(* IEC 61131-3 sources: plc-st-coding-agent/progress/evidence/f14_v6_public_pilot_20261112/jobs/codex_minimax-m27, 42 files *)

(* ---- public-easy-01.candidate_01.st ---- *)
(*
ENGINEERING_CONTRACT
================================================================================
State Machine: Automated Filling Line (5-stage sequential + reset)
Clause ID | Output/State    | Activation          | Retention       | Reset
----------|-----------------|---------------------|-----------------|------------------
PUB003    | Pump_Motor      | bottleSensor=1      | Hold in CLEANING| cleaningConfirmButton (→FILLING)
PUB004    | Filling_Valve   | cleaningConfirmBtn  | Hold in FILLING | fillingConfirmButton (→CAPPING)
PUB005    | Capping_Machine | fillingConfirmBtn   | Hold in CAPPING | cappingConfirmButton (→PACKING)
PUB006    | Packing_Machine | cappingConfirmBtn   | Hold in PACKING | packingConfirmButton (→COMPLETE)
PUB007    | Completion_Light| packingConfirmBtn   | Hold until RESET| finishedButton (→IDLE)
PUB008    | (finishedButton)| Reset all, cycle end| N/A             | Automatic →IDLE
--------------------------------------------------------------------------------
Priority: Same-scan sequential (IDLE→CLEANING→FILLING→CAPPING→PACKING→COMPLETE→IDLE)
Units: None (binary signals, no timeouts specified)
Boundary: bottleSensor rising edge starts CLEANING; finishedButton resets COMPLETE→IDLE
--------------------------------------------------------------------------------
CONTRACT_RULES []
================================================================================
*)

FUNCTION_BLOCK FillingLineControl
VAR_INPUT
    bottleSensor          : BOOL;
    cleaningConfirmButton : BOOL;
    fillingConfirmButton  : BOOL;
    cappingConfirmButton  : BOOL;
    packingConfirmButton  : BOOL;
    finishedButton        : BOOL;
END_VAR
VAR_OUTPUT
    Pump_Motor      : BOOL;
    Filling_Valve   : BOOL;
    Capping_Machine : BOOL;
    Packing_Machine : BOOL;
    Completion_Light: BOOL;
END_VAR
VAR
    eState : INT;
END_VAR

// State enumeration: 0=IDLE, 1=CLEANING, 2=FILLING, 3=CAPPING, 4=PACKING, 5=COMPLETE
CASE eState OF
    0: // IDLE
        Pump_Motor       := FALSE;
        Filling_Valve    := FALSE;
        Capping_Machine  := FALSE;
        Packing_Machine  := FALSE;
        Completion_Light := FALSE;
        IF bottleSensor THEN
            eState := 1; // → CLEANING
        END_IF;

    1: // CLEANING
        Pump_Motor       := TRUE;
        Filling_Valve    := FALSE;
        Capping_Machine  := FALSE;
        Packing_Machine  := FALSE;
        Completion_Light := FALSE;
        IF cleaningConfirmButton THEN
            eState := 2; // → FILLING
        END_IF;

    2: // FILLING
        Pump_Motor       := FALSE;
        Filling_Valve    := TRUE;
        Capping_Machine  := FALSE;
        Packing_Machine  := FALSE;
        Completion_Light := FALSE;
        IF fillingConfirmButton THEN
            eState := 3; // → CAPPING
        END_IF;

    3: // CAPPING
        Pump_Motor       := FALSE;
        Filling_Valve    := FALSE;
        Capping_Machine  := TRUE;
        Packing_Machine  := FALSE;
        Completion_Light := FALSE;
        IF cappingConfirmButton THEN
            eState := 4; // → PACKING
        END_IF;

    4: // PACKING
        Pump_Motor       := FALSE;
        Filling_Valve    := FALSE;
        Capping_Machine  := FALSE;
        Packing_Machine  := TRUE;
        Completion_Light := FALSE;
        IF packingConfirmButton THEN
            eState := 5; // → COMPLETE
        END_IF;

    5: // COMPLETE
        Pump_Motor       := FALSE;
        Filling_Valve    := FALSE;
        Capping_Machine  := FALSE;
        Packing_Machine  := FALSE;
        Completion_Light := TRUE;
        IF finishedButton THEN
            eState := 0; // → IDLE (cycle reset)
        END_IF;

END_CASE;

END_FUNCTION_BLOCK

(* ---- public-easy-01.candidate_02.st ---- *)
(*
ENGINEERING_CONTRACT
================================================================================
State Machine: Automated Filling Line (5-stage sequential + reset)
Clause ID | Output/State    | Activation          | Retention       | Reset
----------|-----------------|---------------------|-----------------|------------------
PUB003    | Pump_Motor      | bottleSensor=1      | Hold in CLEANING| cleaningConfirmButton (→FILLING)
PUB004    | Filling_Valve   | cleaningConfirmBtn  | Hold in FILLING | fillingConfirmButton (→CAPPING)
PUB005    | Capping_Machine | fillingConfirmBtn   | Hold in CAPPING | cappingConfirmButton (→PACKING)
PUB006    | Packing_Machine | cappingConfirmBtn   | Hold in PACKING | packingConfirmButton (→COMPLETE)
PUB007    | Completion_Light| packingConfirmBtn   | Hold until RESET| finishedButton (→IDLE)
PUB008    | (finishedButton)| Reset all, cycle end| N/A             | Automatic →IDLE
--------------------------------------------------------------------------------
Priority: Same-scan sequential (IDLE→CLEANING→FILLING→CAPPING→PACKING→COMPLETE→IDLE)
Units: None (binary signals, no timeouts specified)
Boundary: bottleSensor rising edge starts CLEANING; finishedButton resets COMPLETE→IDLE
--------------------------------------------------------------------------------
CONTRACT_RULES []
================================================================================
*)

FUNCTION_BLOCK FillingLineControl
VAR_INPUT
    bottleSensor          : BOOL;
    cleaningConfirmButton : BOOL;
    fillingConfirmButton  : BOOL;
    cappingConfirmButton  : BOOL;
    packingConfirmButton  : BOOL;
    finishedButton        : BOOL;
END_VAR
VAR_OUTPUT
    Pump_Motor      : BOOL;
    Filling_Valve   : BOOL;
    Capping_Machine : BOOL;
    Packing_Machine : BOOL;
    Completion_Light: BOOL;
END_VAR
VAR
    eState : INT;
END_VAR

// State: 0=IDLE, 1=CLEANING, 2=FILLING, 3=CAPPING, 4=PACKING, 5=COMPLETE
// Multiple transitions within same scan when conditions allow
IF eState = 0 AND bottleSensor THEN
    eState := 1;
END_IF;

IF eState = 1 AND cleaningConfirmButton THEN
    eState := 2;
END_IF;

IF eState = 2 AND fillingConfirmButton THEN
    eState := 3;
END_IF;

IF eState = 3 AND cappingConfirmButton THEN
    eState := 4;
END_IF;

IF eState = 4 AND packingConfirmButton THEN
    eState := 5;
END_IF;

IF eState = 5 AND finishedButton THEN
    eState := 0;
END_IF;

// Output assignment based on current state
IF eState = 1 THEN
    Pump_Motor := TRUE;
END_IF;

IF eState = 2 THEN
    Filling_Valve := TRUE;
END_IF;

IF eState = 3 THEN
    Capping_Machine := TRUE;
END_IF;

IF eState = 4 THEN
    Packing_Machine := TRUE;
END_IF;

IF eState = 5 THEN
    Completion_Light := TRUE;
END_IF;

END_FUNCTION_BLOCK

(* ---- public-easy-01.candidate_03.st ---- *)
(*
ENGINEERING_CONTRACT
================================================================================
State Machine: Automated Filling Line (5-stage sequential + reset)
Clause ID | Output/State    | Activation          | Retention       | Reset
----------|-----------------|---------------------|-----------------|------------------
PUB003    | Pump_Motor      | bottleSensor=1      | Hold in CLEANING| cleaningConfirmButton (→FILLING)
PUB004    | Filling_Valve   | cleaningConfirmBtn  | Hold in FILLING | fillingConfirmButton (→CAPPING)
PUB005    | Capping_Machine | fillingConfirmBtn   | Hold in CAPPING | cappingConfirmButton (→PACKING)
PUB006    | Packing_Machine | cappingConfirmBtn   | Hold in PACKING | packingConfirmButton (→COMPLETE)
PUB007    | Completion_Light| packingConfirmBtn   | Hold until RESET| finishedButton (→IDLE)
PUB008    | (finishedButton)| Reset all, cycle end| N/A             | Automatic →IDLE
--------------------------------------------------------------------------------
Priority: Same-scan sequential (IDLE→CLEANING→FILLING→CAPPING→PACKING→COMPLETE→IDLE)
Units: None (binary signals, no timeouts specified)
Boundary: bottleSensor rising edge starts CLEANING; finishedButton resets COMPLETE→IDLE
--------------------------------------------------------------------------------
CONTRACT_RULES []
================================================================================
*)

FUNCTION_BLOCK FillingLineControl
VAR_INPUT
    bottleSensor          : BOOL;
    cleaningConfirmButton : BOOL;
    fillingConfirmButton  : BOOL;
    cappingConfirmButton  : BOOL;
    packingConfirmButton  : BOOL;
    finishedButton        : BOOL;
END_VAR
VAR_OUTPUT
    Pump_Motor      : BOOL;
    Filling_Valve   : BOOL;
    Capping_Machine : BOOL;
    Packing_Machine : BOOL;
    Completion_Light: BOOL;
END_VAR
VAR
    eState : INT;
END_VAR

// State: 0=IDLE, 1=CLEANING, 2=FILLING, 3=CAPPING, 4=PACKING, 5=COMPLETE
// Reset all outputs each scan to ensure clean state transitions
Pump_Motor      := FALSE;
Filling_Valve   := FALSE;
Capping_Machine := FALSE;
Packing_Machine := FALSE;
Completion_Light:= FALSE;

// State transitions - sequential same-scan processing
IF eState = 0 AND bottleSensor THEN
    eState := 1;
END_IF;

IF eState = 1 AND cleaningConfirmButton THEN
    eState := 2;
END_IF;

IF eState = 2 AND fillingConfirmButton THEN
    eState := 3;
END_IF;

IF eState = 3 AND cappingConfirmButton THEN
    eState := 4;
END_IF;

IF eState = 4 AND packingConfirmButton THEN
    eState := 5;
END_IF;

IF eState = 5 AND finishedButton THEN
    eState := 0;
END_IF;

// Output activation based on current state
IF eState = 1 THEN
    Pump_Motor := TRUE;
END_IF;

IF eState = 2 THEN
    Filling_Valve := TRUE;
END_IF;

IF eState = 3 THEN
    Capping_Machine := TRUE;
END_IF;

IF eState = 4 THEN
    Packing_Machine := TRUE;
END_IF;

IF eState = 5 THEN
    Completion_Light := TRUE;
END_IF;

END_FUNCTION_BLOCK

(* ---- public-easy-01.candidate_04.st ---- *)
Looking at the checkpoint, tc-08 shows ALL outputs TRUE when `finishedButton=true` from a prior state. The issue is that outputs never get reset when transitioning between states—they only get set TRUE but never set FALSE.

(*
ENGINEERING_CONTRACT
================================================================================
State Machine: Automated Filling Line (5-stage sequential + reset)
Clause ID | Output/State    | Activation          | Retention       | Reset
----------|-----------------|---------------------|-----------------|------------------
PUB003    | Pump_Motor      | bottleSensor=1      | Hold in CLEANING| Implicit (output cleared on state exit)
PUB004    | Filling_Valve   | cleaningConfirmBtn  | Hold in FILLING | Implicit (output cleared on state exit)
PUB005    | Capping_Machine | fillingConfirmBtn   | Hold in CAPPING | Implicit (output cleared on state exit)
PUB006    | Packing_Machine | cappingConfirmBtn   | Hold in PACKING | Implicit (output cleared on state exit)
PUB007    | Completion_Light| packingConfirmBtn   | Hold in COMPLETE| Implicit (output cleared on finishedButton reset)
PUB008    | (finishedButton)| Reset all outputs   | N/A             | Automatic →IDLE
--------------------------------------------------------------------------------
Priority: Same-scan sequential (IDLE→CLEANING→FILLING→CAPPING→PACKING→COMPLETE→IDLE)
Units: None (binary signals, no timeouts specified)
Boundary: Outputs are level-based; cleared when state exits, no edge-only behavior
--------------------------------------------------------------------------------
CONTRACT_RULES []
================================================================================
*)

FUNCTION_BLOCK FillingLineControl
VAR_INPUT
    bottleSensor          : BOOL;
    cleaningConfirmButton : BOOL;
    fillingConfirmButton  : BOOL;
    cappingConfirmButton  : BOOL;
    packingConfirmButton  : BOOL;
    finishedButton        : BOOL;
END_VAR
VAR_OUTPUT
    Pump_Motor      : BOOL;
    Filling_Valve   : BOOL;
    Capping_Machine : BOOL;
    Packing_Machine : BOOL;
    Completion_Light: BOOL;
END_VAR
VAR
    eState : INT;
END_VAR

// State: 0=IDLE, 1=CLEANING, 2=FILLING, 3=CAPPING, 4=PACKING, 5=COMPLETE
// Clear all outputs first (no latching across state transitions)
Pump_Motor      := FALSE;
Filling_Valve   := FALSE;
Capping_Machine := FALSE;
Packing_Machine := FALSE;
Completion_Light:= FALSE;

// State transitions (same-scan sequential)
IF eState = 0 AND bottleSensor THEN
    eState := 1;
END_IF;

IF eState = 1 AND cleaningConfirmButton THEN
    eState := 2;
END_IF;

IF eState = 2 AND fillingConfirmButton THEN
    eState := 3;
END_IF;

IF eState = 3 AND cappingConfirmButton THEN
    eState := 4;
END_IF;

IF eState = 4 AND packingConfirmButton THEN
    eState := 5;
END_IF;

IF eState = 5 AND finishedButton THEN
    eState := 0;
END_IF;

// Output assignment based on current state (level-based, cleared on exit)
IF eState = 1 THEN
    Pump_Motor := TRUE;
END_IF;

IF eState = 2 THEN
    Filling_Valve := TRUE;
END_IF;

IF eState = 3 THEN
    Capping_Machine := TRUE;
END_IF;

IF eState = 4 THEN
    Packing_Machine := TRUE;
END_IF;

IF eState = 5 THEN
    Completion_Light := TRUE;
END_IF;

END_FUNCTION_BLOCK

(* ---- public-easy-01.raw_candidate_01.st ---- *)
(*
ENGINEERING_CONTRACT
================================================================================
State Machine: Automated Filling Line (5-stage sequential + reset)
Clause ID | Output/State    | Activation          | Retention       | Reset
----------|-----------------|---------------------|-----------------|------------------
PUB003    | Pump_Motor      | bottleSensor=1      | Hold in CLEANING| cleaningConfirmButton (→FILLING)
PUB004    | Filling_Valve   | cleaningConfirmBtn  | Hold in FILLING | fillingConfirmButton (→CAPPING)
PUB005    | Capping_Machine | fillingConfirmBtn   | Hold in CAPPING | cappingConfirmButton (→PACKING)
PUB006    | Packing_Machine | cappingConfirmBtn   | Hold in PACKING | packingConfirmButton (→COMPLETE)
PUB007    | Completion_Light| packingConfirmBtn   | Hold until RESET| finishedButton (→IDLE)
PUB008    | (finishedButton)| Reset all, cycle end| N/A             | Automatic →IDLE
--------------------------------------------------------------------------------
Priority: Same-scan sequential (IDLE→CLEANING→FILLING→CAPPING→PACKING→COMPLETE→IDLE)
Units: None (binary signals, no timeouts specified)
Boundary: bottleSensor rising edge starts CLEANING; finishedButton resets COMPLETE→IDLE
--------------------------------------------------------------------------------
CONTRACT_RULES []
================================================================================
*)

FUNCTION_BLOCK FillingLineControl
VAR_INPUT
    bottleSensor          : BOOL;
    cleaningConfirmButton : BOOL;
    fillingConfirmButton  : BOOL;
    cappingConfirmButton  : BOOL;
    packingConfirmButton  : BOOL;
    finishedButton        : BOOL;
END_VAR
VAR_OUTPUT
    Pump_Motor      : BOOL;
    Filling_Valve   : BOOL;
    Capping_Machine : BOOL;
    Packing_Machine : BOOL;
    Completion_Light: BOOL;
END_VAR
VAR
    eState : INT;
END_VAR

// State enumeration: 0=IDLE, 1=CLEANING, 2=FILLING, 3=CAPPING, 4=PACKING, 5=COMPLETE
CASE eState OF
    0: // IDLE
        Pump_Motor       := FALSE;
        Filling_Valve    := FALSE;
        Capping_Machine  := FALSE;
        Packing_Machine  := FALSE;
        Completion_Light := FALSE;
        IF bottleSensor THEN
            eState := 1; // → CLEANING
        END_IF;

    1: // CLEANING
        Pump_Motor       := TRUE;
        Filling_Valve    := FALSE;
        Capping_Machine  := FALSE;
        Packing_Machine  := FALSE;
        Completion_Light := FALSE;
        IF cleaningConfirmButton THEN
            eState := 2; // → FILLING
        END_IF;

    2: // FILLING
        Pump_Motor       := FALSE;
        Filling_Valve    := TRUE;
        Capping_Machine  := FALSE;
        Packing_Machine  := FALSE;
        Completion_Light := FALSE;
        IF fillingConfirmButton THEN
            eState := 3; // → CAPPING
        END_IF;

    3: // CAPPING
        Pump_Motor       := FALSE;
        Filling_Valve    := FALSE;
        Capping_Machine  := TRUE;
        Packing_Machine  := FALSE;
        Completion_Light := FALSE;
        IF cappingConfirmButton THEN
            eState := 4; // → PACKING
        END_IF;

    4: // PACKING
        Pump_Motor       := FALSE;
        Filling_Valve    := FALSE;
        Capping_Machine  := FALSE;
        Packing_Machine  := TRUE;
        Completion_Light := FALSE;
        IF packingConfirmButton THEN
            eState := 5; // → COMPLETE
        END_IF;

    5: // COMPLETE
        Pump_Motor       := FALSE;
        Filling_Valve    := FALSE;
        Capping_Machine  := FALSE;
        Packing_Machine  := FALSE;
        Completion_Light := TRUE;
        IF finishedButton THEN
            eState := 0; // → IDLE (cycle reset)
        END_IF;

END_CASE;

END_FUNCTION_BLOCK

(* ---- public-easy-01.raw_candidate_02.st ---- *)
(*
ENGINEERING_CONTRACT
================================================================================
State Machine: Automated Filling Line (5-stage sequential + reset)
Clause ID | Output/State    | Activation          | Retention       | Reset
----------|-----------------|---------------------|-----------------|------------------
PUB003    | Pump_Motor      | bottleSensor=1      | Hold in CLEANING| cleaningConfirmButton (→FILLING)
PUB004    | Filling_Valve   | cleaningConfirmBtn  | Hold in FILLING | fillingConfirmButton (→CAPPING)
PUB005    | Capping_Machine | fillingConfirmBtn   | Hold in CAPPING | cappingConfirmButton (→PACKING)
PUB006    | Packing_Machine | cappingConfirmBtn   | Hold in PACKING | packingConfirmButton (→COMPLETE)
PUB007    | Completion_Light| packingConfirmBtn   | Hold until RESET| finishedButton (→IDLE)
PUB008    | (finishedButton)| Reset all, cycle end| N/A             | Automatic →IDLE
--------------------------------------------------------------------------------
Priority: Same-scan sequential (IDLE→CLEANING→FILLING→CAPPING→PACKING→COMPLETE→IDLE)
Units: None (binary signals, no timeouts specified)
Boundary: bottleSensor rising edge starts CLEANING; finishedButton resets COMPLETE→IDLE
--------------------------------------------------------------------------------
CONTRACT_RULES []
================================================================================
*)

FUNCTION_BLOCK FillingLineControl
VAR_INPUT
    bottleSensor          : BOOL;
    cleaningConfirmButton : BOOL;
    fillingConfirmButton  : BOOL;
    cappingConfirmButton  : BOOL;
    packingConfirmButton  : BOOL;
    finishedButton        : BOOL;
END_VAR
VAR_OUTPUT
    Pump_Motor      : BOOL;
    Filling_Valve   : BOOL;
    Capping_Machine : BOOL;
    Packing_Machine : BOOL;
    Completion_Light: BOOL;
END_VAR
VAR
    eState : INT;
END_VAR

// State: 0=IDLE, 1=CLEANING, 2=FILLING, 3=CAPPING, 4=PACKING, 5=COMPLETE
// Multiple transitions within same scan when conditions allow
IF eState = 0 AND bottleSensor THEN
    eState := 1;
END_IF;

IF eState = 1 AND cleaningConfirmButton THEN
    eState := 2;
END_IF;

IF eState = 2 AND fillingConfirmButton THEN
    eState := 3;
END_IF;

IF eState = 3 AND cappingConfirmButton THEN
    eState := 4;
END_IF;

IF eState = 4 AND packingConfirmButton THEN
    eState := 5;
END_IF;

IF eState = 5 AND finishedButton THEN
    eState := 0;
END_IF;

// Output assignment based on current state
IF eState = 1 THEN
    Pump_Motor := TRUE;
END_IF;

IF eState = 2 THEN
    Filling_Valve := TRUE;
END_IF;

IF eState = 3 THEN
    Capping_Machine := TRUE;
END_IF;

IF eState = 4 THEN
    Packing_Machine := TRUE;
END_IF;

IF eState = 5 THEN
    Completion_Light := TRUE;
END_IF;

END_FUNCTION_BLOCK

(* ---- public-easy-01.raw_candidate_03.st ---- *)
(*
ENGINEERING_CONTRACT
================================================================================
State Machine: Automated Filling Line (5-stage sequential + reset)
Clause ID | Output/State    | Activation          | Retention       | Reset
----------|-----------------|---------------------|-----------------|------------------
PUB003    | Pump_Motor      | bottleSensor=1      | Hold in CLEANING| cleaningConfirmButton (→FILLING)
PUB004    | Filling_Valve   | cleaningConfirmBtn  | Hold in FILLING | fillingConfirmButton (→CAPPING)
PUB005    | Capping_Machine | fillingConfirmBtn   | Hold in CAPPING | cappingConfirmButton (→PACKING)
PUB006    | Packing_Machine | cappingConfirmBtn   | Hold in PACKING | packingConfirmButton (→COMPLETE)
PUB007    | Completion_Light| packingConfirmBtn   | Hold until RESET| finishedButton (→IDLE)
PUB008    | (finishedButton)| Reset all, cycle end| N/A             | Automatic →IDLE
--------------------------------------------------------------------------------
Priority: Same-scan sequential (IDLE→CLEANING→FILLING→CAPPING→PACKING→COMPLETE→IDLE)
Units: None (binary signals, no timeouts specified)
Boundary: bottleSensor rising edge starts CLEANING; finishedButton resets COMPLETE→IDLE
--------------------------------------------------------------------------------
CONTRACT_RULES []
================================================================================
*)

FUNCTION_BLOCK FillingLineControl
VAR_INPUT
    bottleSensor          : BOOL;
    cleaningConfirmButton : BOOL;
    fillingConfirmButton  : BOOL;
    cappingConfirmButton  : BOOL;
    packingConfirmButton  : BOOL;
    finishedButton        : BOOL;
END_VAR
VAR_OUTPUT
    Pump_Motor      : BOOL;
    Filling_Valve   : BOOL;
    Capping_Machine : BOOL;
    Packing_Machine : BOOL;
    Completion_Light: BOOL;
END_VAR
VAR
    eState : INT;
END_VAR

// State: 0=IDLE, 1=CLEANING, 2=FILLING, 3=CAPPING, 4=PACKING, 5=COMPLETE
// Reset all outputs each scan to ensure clean state transitions
Pump_Motor      := FALSE;
Filling_Valve   := FALSE;
Capping_Machine := FALSE;
Packing_Machine := FALSE;
Completion_Light:= FALSE;

// State transitions - sequential same-scan processing
IF eState = 0 AND bottleSensor THEN
    eState := 1;
END_IF;

IF eState = 1 AND cleaningConfirmButton THEN
    eState := 2;
END_IF;

IF eState = 2 AND fillingConfirmButton THEN
    eState := 3;
END_IF;

IF eState = 3 AND cappingConfirmButton THEN
    eState := 4;
END_IF;

IF eState = 4 AND packingConfirmButton THEN
    eState := 5;
END_IF;

IF eState = 5 AND finishedButton THEN
    eState := 0;
END_IF;

// Output activation based on current state
IF eState = 1 THEN
    Pump_Motor := TRUE;
END_IF;

IF eState = 2 THEN
    Filling_Valve := TRUE;
END_IF;

IF eState = 3 THEN
    Capping_Machine := TRUE;
END_IF;

IF eState = 4 THEN
    Packing_Machine := TRUE;
END_IF;

IF eState = 5 THEN
    Completion_Light := TRUE;
END_IF;

END_FUNCTION_BLOCK

(* ---- public-easy-01.raw_candidate_04.st ---- *)
Looking at the checkpoint, tc-08 shows ALL outputs TRUE when `finishedButton=true` from a prior state. The issue is that outputs never get reset when transitioning between states—they only get set TRUE but never set FALSE.

(*
ENGINEERING_CONTRACT
================================================================================
State Machine: Automated Filling Line (5-stage sequential + reset)
Clause ID | Output/State    | Activation          | Retention       | Reset
----------|-----------------|---------------------|-----------------|------------------
PUB003    | Pump_Motor      | bottleSensor=1      | Hold in CLEANING| Implicit (output cleared on state exit)
PUB004    | Filling_Valve   | cleaningConfirmBtn  | Hold in FILLING | Implicit (output cleared on state exit)
PUB005    | Capping_Machine | fillingConfirmBtn   | Hold in CAPPING | Implicit (output cleared on state exit)
PUB006    | Packing_Machine | cappingConfirmBtn   | Hold in PACKING | Implicit (output cleared on state exit)
PUB007    | Completion_Light| packingConfirmBtn   | Hold in COMPLETE| Implicit (output cleared on finishedButton reset)
PUB008    | (finishedButton)| Reset all outputs   | N/A             | Automatic →IDLE
--------------------------------------------------------------------------------
Priority: Same-scan sequential (IDLE→CLEANING→FILLING→CAPPING→PACKING→COMPLETE→IDLE)
Units: None (binary signals, no timeouts specified)
Boundary: Outputs are level-based; cleared when state exits, no edge-only behavior
--------------------------------------------------------------------------------
CONTRACT_RULES []
================================================================================
*)

FUNCTION_BLOCK FillingLineControl
VAR_INPUT
    bottleSensor          : BOOL;
    cleaningConfirmButton : BOOL;
    fillingConfirmButton  : BOOL;
    cappingConfirmButton  : BOOL;
    packingConfirmButton  : BOOL;
    finishedButton        : BOOL;
END_VAR
VAR_OUTPUT
    Pump_Motor      : BOOL;
    Filling_Valve   : BOOL;
    Capping_Machine : BOOL;
    Packing_Machine : BOOL;
    Completion_Light: BOOL;
END_VAR
VAR
    eState : INT;
END_VAR

// State: 0=IDLE, 1=CLEANING, 2=FILLING, 3=CAPPING, 4=PACKING, 5=COMPLETE
// Clear all outputs first (no latching across state transitions)
Pump_Motor      := FALSE;
Filling_Valve   := FALSE;
Capping_Machine := FALSE;
Packing_Machine := FALSE;
Completion_Light:= FALSE;

// State transitions (same-scan sequential)
IF eState = 0 AND bottleSensor THEN
    eState := 1;
END_IF;

IF eState = 1 AND cleaningConfirmButton THEN
    eState := 2;
END_IF;

IF eState = 2 AND fillingConfirmButton THEN
    eState := 3;
END_IF;

IF eState = 3 AND cappingConfirmButton THEN
    eState := 4;
END_IF;

IF eState = 4 AND packingConfirmButton THEN
    eState := 5;
END_IF;

IF eState = 5 AND finishedButton THEN
    eState := 0;
END_IF;

// Output assignment based on current state (level-based, cleared on exit)
IF eState = 1 THEN
    Pump_Motor := TRUE;
END_IF;

IF eState = 2 THEN
    Filling_Valve := TRUE;
END_IF;

IF eState = 3 THEN
    Capping_Machine := TRUE;
END_IF;

IF eState = 4 THEN
    Packing_Machine := TRUE;
END_IF;

IF eState = 5 THEN
    Completion_Light := TRUE;
END_IF;

END_FUNCTION_BLOCK

(* ---- public-easy-04.candidate_01.st ---- *)
(*
ENGINEERING_CONTRACT
===================
PUB001: Jam transfer pump control - viscosity debouncing, E-stop, runtime, maintenance

Output States:
- VFD_RUN:
  - Activation: TRUE when PASTE_E_STOP_NC=TRUE AND viscosity_valid=TRUE
  - Retention: Hold TRUE across scans while conditions remain valid
  - Explicit Reset: Immediate OFF on PASTE_E_STOP_NC=FALSE
  - Same-scan Priority: Evaluated after safety check (E-stop wins)

- PUMP_RUNTIME_ACC:
  - Activation: Increments by CycleTime each scan when VFD_RUN=TRUE
  - Retention: Maintains value when VFD_RUN=FALSE (no decay)
  - Reset: Zero at power-up only (PUB006)
  - Units: LTIME (nanoseconds)

- PUMP_MAINT_DUE:
  - Activation: Set TRUE when PUMP_RUNTIME_ACC >= 500 hours
  - Retention: Hold TRUE once set (informational, PUB005)
  - Reset: Not specified (no auto-reset)
  - Units: LTIME comparison vs 500*3600*1e9 nanoseconds

Safety:
- E-stop (PASTE_E_STOP_NC=FALSE) immediately disables VFD_RUN
- E-stop clears any incomplete debounce timing (TON disabled resets)
- Maintenance indication does not affect pump operation or safety (PUB005)
*)

(* CONTRACT_RULES [] *)

FUNCTION_BLOCK JamPumpControl
VAR_INPUT
    VISCOSITY_OK    : BOOL;
    PASTE_E_STOP_NC : BOOL;
    DebounceTime    : TIME;
    CycleTime       : TIME;
END_VAR

VAR_OUTPUT
    VFD_RUN         : BOOL;
    PUMP_MAINT_DUE  : BOOL;
    PUMP_RUNTIME_ACC: LTIME;
END_VAR

VAR
    ViscosityDebounce : TON;
    tmpViscosityValid : BOOL;
END_VAR

tmpViscosityValid := ViscosityDebounce.Q;

IF NOT PASTE_E_STOP_NC THEN
    VFD_RUN := FALSE;
    ViscosityDebounce(IN := FALSE, PT := DebounceTime);
    tmpViscosityValid := FALSE;
ELSIF VISCOSITY_OK THEN
    ViscosityDebounce(IN := TRUE, PT := DebounceTime);
ELSE
    ViscosityDebounce(IN := FALSE, PT := DebounceTime);
    tmpViscosityValid := FALSE;
END_IF;

IF PASTE_E_STOP_NC AND tmpViscosityValid THEN
    VFD_RUN := TRUE;
ELSE
    VFD_RUN := FALSE;
END_IF;

IF VFD_RUN THEN
    PUMP_RUNTIME_ACC := PUMP_RUNTIME_ACC + TO_LTIME(CycleTime);
END_IF;

IF PUMP_RUNTIME_ACC >= TO_LTIME(TIME_TO_LTIME(T#500h)) THEN
    PUMP_MAINT_DUE := TRUE;
END_IF;

ViscosityDebounce(IN := ViscosityDebounce.IN, PT := DebounceTime);

END_FUNCTION_BLOCK

(* ---- public-easy-04.candidate_02.st ---- *)
(*
ENGINEERING_CONTRACT
===================
PUB001: Jam transfer pump control - viscosity debouncing, E-stop, runtime, maintenance

Output States (Pub Clause IDs):
- VFD_RUN (PUB002, PUB003):
  - Activation: TRUE when PASTE_E_STOP_NC=TRUE AND viscosity_valid=TRUE (debounce complete)
  - Retention: Hold TRUE across scans while conditions remain valid
  - Explicit Reset: Immediate OFF when PASTE_E_STOP_NC=FALSE (PUB003), also OFF when viscosity invalidates
  - Same-scan Priority: Safety check (E-stop) evaluated first; viscosity check completes debounce timing

- PUMP_RUNTIME_ACC (PUB004):
  - Activation: Increments by CycleTime*1e6 (ms to ns) each scan when VFD_RUN=TRUE
  - Retention: Maintains value when VFD_RUN=FALSE (no decay, PUB004 preserved across stops)
  - Reset: Zero at power-up only (PUB006); no auto-reset during operation
  - Units: LTIME nanoseconds; 500 hours = 1.8e12 ns for comparison

- PUMP_MAINT_DUE (PUB005):
  - Activation: Set TRUE when PUMP_RUNTIME_ACC >= 500 hours (LTIME#500h in ns)
  - Retention: Hold TRUE once set (informational, PUB005 specifies no auto-reset requirement)
  - Reset: Not specified; no reset implemented
  - Units: LTIME nanoseconds, 500 hours = 500*3600*1e9 = 1.8e12 nanoseconds

Safety (PUB003):
- E-stop (PASTE_E_STOP_NC=FALSE) immediately disables VFD_RUN
- E-stop clears any incomplete debounce timing (TON disabled via IN=FALSE resets ET to 0)
- Maintenance indication does not affect pump operation or safety (PUB005)
*)

(* CONTRACT_RULES [] *)

FUNCTION_BLOCK JamPumpControl
VAR_INPUT
    VISCOSITY_OK    : BOOL;
    PASTE_E_STOP_NC : BOOL;
    DebounceTime    : TIME;
    CycleTime       : TIME;
END_VAR

VAR_OUTPUT
    VFD_RUN         : BOOL;
    PUMP_MAINT_DUE  : BOOL;
    PUMP_RUNTIME_ACC: LTIME;
END_VAR

VAR
    ViscosityDebounce : TON;
    tmpViscosityValid : BOOL;
    tmpLocalIN        : BOOL;
END_VAR

IF NOT PASTE_E_STOP_NC THEN
    tmpLocalIN := FALSE;
ELSIF VISCOSITY_OK THEN
    tmpLocalIN := TRUE;
ELSE
    tmpLocalIN := FALSE;
END_IF;

ViscosityDebounce(IN := tmpLocalIN, PT := DebounceTime);
tmpViscosityValid := ViscosityDebounce.Q;

IF PASTE_E_STOP_NC AND tmpViscosityValid THEN
    VFD_RUN := TRUE;
ELSE
    VFD_RUN := FALSE;
END_IF;

IF VFD_RUN THEN
    PUMP_RUNTIME_ACC := PUMP_RUNTIME_ACC + TO_LTIME(CycleTime) * 1000000;
END_IF;

IF PUMP_RUNTIME_ACC >= TO_LTIME(T#500h) THEN
    PUMP_MAINT_DUE := TRUE;
END_IF;

END_FUNCTION_BLOCK

(* ---- public-easy-04.candidate_03.st ---- *)
(*
ENGINEERING_CONTRACT
===================
PUB001: Jam transfer pump control - viscosity debouncing, E-stop, runtime, maintenance

Output States:
- VFD_RUN:
  - Activation: TRUE when PASTE_E_STOP_NC=TRUE AND viscosity_valid=TRUE (TON.Q)
  - Retention: Hold TRUE across scans while conditions remain valid
  - Explicit Reset: Immediate OFF on PASTE_E_STOP_NC=FALSE (PUB003)
  - Same-scan Priority: E-stop disables first, then viscosity checked
  - Units: Boolean permissive

- PUMP_RUNTIME_ACC:
  - Activation: Increment by CycleTime each scan when VFD_RUN=TRUE (PUB004)
  - Retention: Maintains value when VFD_RUN=FALSE (no decay)
  - Reset: Zero at power-up only (PUB006)
  - Units: LTIME nanoseconds

- PUMP_MAINT_DUE:
  - Activation: Set TRUE when PUMP_RUNTIME_ACC >= 500 hours (PUB005)
  - Retention: Hold TRUE once set (informational, no auto-reset per PUB005)
  - Reset: Not specified
  - Units: LTIME comparison

Safety:
- E-stop (PASTE_E_STOP_NC=FALSE) immediately disables VFD_RUN (PUB003)
- E-stop clears debounce by disabling TON (PUB003)
- Maintenance has no effect on operation or safety (PUB005)
*)

(* CONTRACT_RULES [] *)

FUNCTION_BLOCK JamPumpControl
VAR_INPUT
    VISCOSITY_OK    : BOOL;
    PASTE_E_STOP_NC : BOOL;
    DebounceTime    : TIME;
    CycleTime       : TIME;
END_VAR

VAR_OUTPUT
    VFD_RUN         : BOOL;
    PUMP_MAINT_DUE  : BOOL;
    PUMP_RUNTIME_ACC: LTIME;
END_VAR

VAR
    ViscosityDebounce : TON;
END_VAR

ViscosityDebounce(
    IN  := PASTE_E_STOP_NC AND VISCOSITY_OK,
    PT  := DebounceTime
);

VFD_RUN := PASTE_E_STOP_NC AND ViscosityDebounce.Q;

IF VFD_RUN THEN
    PUMP_RUNTIME_ACC := PUMP_RUNTIME_ACC + TO_LTIME(CycleTime);
END_IF;

IF PUMP_RUNTIME_ACC >= T#500h THEN
    PUMP_MAINT_DUE := TRUE;
END_IF;

END_FUNCTION_BLOCK

(* ---- public-easy-04.candidate_04.st ---- *)
(*
ENGINEERING_CONTRACT
===================
PUB001: Jam transfer pump control - viscosity debouncing, E-stop, runtime, maintenance

Output States:
- VFD_RUN:
  - Activation: TRUE when PASTE_E_STOP_NC=TRUE AND viscosity_valid=TRUE
  - Retention: Hold TRUE across scans while conditions remain valid
  - Explicit Reset: Immediate OFF on PASTE_E_STOP_NC=FALSE
  - Same-scan Priority: Evaluated after safety check (E-stop wins)

- PUMP_RUNTIME_ACC:
  - Activation: Increments by CycleTime each scan when VFD_RUN=TRUE
  - Retention: Maintains value when VFD_RUN=FALSE (no decay)
  - Reset: Zero at power-up only (PUB006)
  - Units: LTIME (nanoseconds)

- PUMP_MAINT_DUE:
  - Activation: Set TRUE when PUMP_RUNTIME_ACC >= 500 hours
  - Retention: Hold TRUE once set (informational, PUB005)
  - Reset: Not specified (no auto-reset)
  - Units: LTIME comparison vs 500*3600*1e9 nanoseconds

Safety:
- E-stop (PASTE_E_STOP_NC=FALSE) immediately disables VFD_RUN
- E-stop clears any incomplete debounce timing (TON disabled resets)
- Maintenance indication does not affect pump operation or safety (PUB005)
*)

(* CONTRACT_RULES [] *)

FUNCTION_BLOCK JamPumpControl
VAR_INPUT
    VISCOSITY_OK    : BOOL;
    PASTE_E_STOP_NC : BOOL;
    DebounceTime    : TIME;
    CycleTime       : TIME;
END_VAR

VAR_OUTPUT
    VFD_RUN         : BOOL;
    PUMP_MAINT_DUE  : BOOL;
    PUMP_RUNTIME_ACC: LTIME;
END_VAR

VAR
    ViscosityDebounce : TON;
    tmpViscosityValid : BOOL;
END_VAR

// Single TON call per scan with correct input determined by E-stop
IF NOT PASTE_E_STOP_NC THEN
    ViscosityDebounce(IN := FALSE, PT := DebounceTime);
ELSE
    ViscosityDebounce(IN := VISCOSITY_OK, PT := DebounceTime);
END_IF;

tmpViscosityValid := ViscosityDebounce.Q;

IF NOT PASTE_E_STOP_NC THEN
    VFD_RUN := FALSE;
ELSE
    VFD_RUN := tmpViscosityValid;
END_IF;

IF VFD_RUN THEN
    PUMP_RUNTIME_ACC := PUMP_RUNTIME_ACC + TO_LTIME(CycleTime);
END_IF;

IF PUMP_RUNTIME_ACC >= T#500h THEN
    PUMP_MAINT_DUE := TRUE;
END_IF;

END_FUNCTION_BLOCK

(* ---- public-easy-04.raw_candidate_01.st ---- *)
(*
ENGINEERING_CONTRACT
===================
PUB001: Jam transfer pump control - viscosity debouncing, E-stop, runtime, maintenance

Output States:
- VFD_RUN:
  - Activation: TRUE when PASTE_E_STOP_NC=TRUE AND viscosity_valid=TRUE
  - Retention: Hold TRUE across scans while conditions remain valid
  - Explicit Reset: Immediate OFF on PASTE_E_STOP_NC=FALSE
  - Same-scan Priority: Evaluated after safety check (E-stop wins)

- PUMP_RUNTIME_ACC:
  - Activation: Increments by CycleTime each scan when VFD_RUN=TRUE
  - Retention: Maintains value when VFD_RUN=FALSE (no decay)
  - Reset: Zero at power-up only (PUB006)
  - Units: LTIME (nanoseconds)

- PUMP_MAINT_DUE:
  - Activation: Set TRUE when PUMP_RUNTIME_ACC >= 500 hours
  - Retention: Hold TRUE once set (informational, PUB005)
  - Reset: Not specified (no auto-reset)
  - Units: LTIME comparison vs 500*3600*1e9 nanoseconds

Safety:
- E-stop (PASTE_E_STOP_NC=FALSE) immediately disables VFD_RUN
- E-stop clears any incomplete debounce timing (TON disabled resets)
- Maintenance indication does not affect pump operation or safety (PUB005)
*)

(* CONTRACT_RULES [] *)

FUNCTION_BLOCK JamPumpControl
VAR_INPUT
    VISCOSITY_OK    : BOOL;
    PASTE_E_STOP_NC : BOOL;
    DebounceTime    : TIME;
    CycleTime       : TIME;
END_VAR

VAR_OUTPUT
    VFD_RUN         : BOOL;
    PUMP_MAINT_DUE  : BOOL;
    PUMP_RUNTIME_ACC: LTIME;
END_VAR

VAR
    ViscosityDebounce : TON;
    tmpViscosityValid : BOOL;
END_VAR

tmpViscosityValid := ViscosityDebounce.Q;

IF NOT PASTE_E_STOP_NC THEN
    VFD_RUN := FALSE;
    ViscosityDebounce(IN := FALSE, PT := DebounceTime);
    tmpViscosityValid := FALSE;
ELSIF VISCOSITY_OK THEN
    ViscosityDebounce(IN := TRUE, PT := DebounceTime);
ELSE
    ViscosityDebounce(IN := FALSE, PT := DebounceTime);
    tmpViscosityValid := FALSE;
END_IF;

IF PASTE_E_STOP_NC AND tmpViscosityValid THEN
    VFD_RUN := TRUE;
ELSE
    VFD_RUN := FALSE;
END_IF;

IF VFD_RUN THEN
    PUMP_RUNTIME_ACC := PUMP_RUNTIME_ACC + TO_LTIME(CycleTime);
END_IF;

IF PUMP_RUNTIME_ACC >= TO_LTIME(TIME_TO_LTIME(T#500h)) THEN
    PUMP_MAINT_DUE := TRUE;
END_IF;

ViscosityDebounce(IN := ViscosityDebounce.IN, PT := DebounceTime);

END_FUNCTION_BLOCK

(* ---- public-easy-04.raw_candidate_02.st ---- *)
(*
ENGINEERING_CONTRACT
===================
PUB001: Jam transfer pump control - viscosity debouncing, E-stop, runtime, maintenance

Output States (Pub Clause IDs):
- VFD_RUN (PUB002, PUB003):
  - Activation: TRUE when PASTE_E_STOP_NC=TRUE AND viscosity_valid=TRUE (debounce complete)
  - Retention: Hold TRUE across scans while conditions remain valid
  - Explicit Reset: Immediate OFF when PASTE_E_STOP_NC=FALSE (PUB003), also OFF when viscosity invalidates
  - Same-scan Priority: Safety check (E-stop) evaluated first; viscosity check completes debounce timing

- PUMP_RUNTIME_ACC (PUB004):
  - Activation: Increments by CycleTime*1e6 (ms to ns) each scan when VFD_RUN=TRUE
  - Retention: Maintains value when VFD_RUN=FALSE (no decay, PUB004 preserved across stops)
  - Reset: Zero at power-up only (PUB006); no auto-reset during operation
  - Units: LTIME nanoseconds; 500 hours = 1.8e12 ns for comparison

- PUMP_MAINT_DUE (PUB005):
  - Activation: Set TRUE when PUMP_RUNTIME_ACC >= 500 hours (LTIME#500h in ns)
  - Retention: Hold TRUE once set (informational, PUB005 specifies no auto-reset requirement)
  - Reset: Not specified; no reset implemented
  - Units: LTIME nanoseconds, 500 hours = 500*3600*1e9 = 1.8e12 nanoseconds

Safety (PUB003):
- E-stop (PASTE_E_STOP_NC=FALSE) immediately disables VFD_RUN
- E-stop clears any incomplete debounce timing (TON disabled via IN=FALSE resets ET to 0)
- Maintenance indication does not affect pump operation or safety (PUB005)
*)

(* CONTRACT_RULES [] *)

FUNCTION_BLOCK JamPumpControl
VAR_INPUT
    VISCOSITY_OK    : BOOL;
    PASTE_E_STOP_NC : BOOL;
    DebounceTime    : TIME;
    CycleTime       : TIME;
END_VAR

VAR_OUTPUT
    VFD_RUN         : BOOL;
    PUMP_MAINT_DUE  : BOOL;
    PUMP_RUNTIME_ACC: LTIME;
END_VAR

VAR
    ViscosityDebounce : TON;
    tmpViscosityValid : BOOL;
    tmpLocalIN        : BOOL;
END_VAR

IF NOT PASTE_E_STOP_NC THEN
    tmpLocalIN := FALSE;
ELSIF VISCOSITY_OK THEN
    tmpLocalIN := TRUE;
ELSE
    tmpLocalIN := FALSE;
END_IF;

ViscosityDebounce(IN := tmpLocalIN, PT := DebounceTime);
tmpViscosityValid := ViscosityDebounce.Q;

IF PASTE_E_STOP_NC AND tmpViscosityValid THEN
    VFD_RUN := TRUE;
ELSE
    VFD_RUN := FALSE;
END_IF;

IF VFD_RUN THEN
    PUMP_RUNTIME_ACC := PUMP_RUNTIME_ACC + TO_LTIME(CycleTime) * 1000000;
END_IF;

IF PUMP_RUNTIME_ACC >= TO_LTIME(T#500h) THEN
    PUMP_MAINT_DUE := TRUE;
END_IF;

END_FUNCTION_BLOCK

(* ---- public-easy-04.raw_candidate_03.st ---- *)
(*
ENGINEERING_CONTRACT
===================
PUB001: Jam transfer pump control - viscosity debouncing, E-stop, runtime, maintenance

Output States:
- VFD_RUN:
  - Activation: TRUE when PASTE_E_STOP_NC=TRUE AND viscosity_valid=TRUE (TON.Q)
  - Retention: Hold TRUE across scans while conditions remain valid
  - Explicit Reset: Immediate OFF on PASTE_E_STOP_NC=FALSE (PUB003)
  - Same-scan Priority: E-stop disables first, then viscosity checked
  - Units: Boolean permissive

- PUMP_RUNTIME_ACC:
  - Activation: Increment by CycleTime each scan when VFD_RUN=TRUE (PUB004)
  - Retention: Maintains value when VFD_RUN=FALSE (no decay)
  - Reset: Zero at power-up only (PUB006)
  - Units: LTIME nanoseconds

- PUMP_MAINT_DUE:
  - Activation: Set TRUE when PUMP_RUNTIME_ACC >= 500 hours (PUB005)
  - Retention: Hold TRUE once set (informational, no auto-reset per PUB005)
  - Reset: Not specified
  - Units: LTIME comparison

Safety:
- E-stop (PASTE_E_STOP_NC=FALSE) immediately disables VFD_RUN (PUB003)
- E-stop clears debounce by disabling TON (PUB003)
- Maintenance has no effect on operation or safety (PUB005)
*)

(* CONTRACT_RULES [] *)

FUNCTION_BLOCK JamPumpControl
VAR_INPUT
    VISCOSITY_OK    : BOOL;
    PASTE_E_STOP_NC : BOOL;
    DebounceTime    : TIME;
    CycleTime       : TIME;
END_VAR

VAR_OUTPUT
    VFD_RUN         : BOOL;
    PUMP_MAINT_DUE  : BOOL;
    PUMP_RUNTIME_ACC: LTIME;
END_VAR

VAR
    ViscosityDebounce : TON;
END_VAR

ViscosityDebounce(
    IN  := PASTE_E_STOP_NC AND VISCOSITY_OK,
    PT  := DebounceTime
);

VFD_RUN := PASTE_E_STOP_NC AND ViscosityDebounce.Q;

IF VFD_RUN THEN
    PUMP_RUNTIME_ACC := PUMP_RUNTIME_ACC + TO_LTIME(CycleTime);
END_IF;

IF PUMP_RUNTIME_ACC >= T#500h THEN
    PUMP_MAINT_DUE := TRUE;
END_IF;

END_FUNCTION_BLOCK

(* ---- public-easy-04.raw_candidate_04.st ---- *)
(*
ENGINEERING_CONTRACT
===================
PUB001: Jam transfer pump control - viscosity debouncing, E-stop, runtime, maintenance

Output States:
- VFD_RUN:
  - Activation: TRUE when PASTE_E_STOP_NC=TRUE AND viscosity_valid=TRUE
  - Retention: Hold TRUE across scans while conditions remain valid
  - Explicit Reset: Immediate OFF on PASTE_E_STOP_NC=FALSE
  - Same-scan Priority: Evaluated after safety check (E-stop wins)

- PUMP_RUNTIME_ACC:
  - Activation: Increments by CycleTime each scan when VFD_RUN=TRUE
  - Retention: Maintains value when VFD_RUN=FALSE (no decay)
  - Reset: Zero at power-up only (PUB006)
  - Units: LTIME (nanoseconds)

- PUMP_MAINT_DUE:
  - Activation: Set TRUE when PUMP_RUNTIME_ACC >= 500 hours
  - Retention: Hold TRUE once set (informational, PUB005)
  - Reset: Not specified (no auto-reset)
  - Units: LTIME comparison vs 500*3600*1e9 nanoseconds

Safety:
- E-stop (PASTE_E_STOP_NC=FALSE) immediately disables VFD_RUN
- E-stop clears any incomplete debounce timing (TON disabled resets)
- Maintenance indication does not affect pump operation or safety (PUB005)
*)

(* CONTRACT_RULES [] *)

FUNCTION_BLOCK JamPumpControl
VAR_INPUT
    VISCOSITY_OK    : BOOL;
    PASTE_E_STOP_NC : BOOL;
    DebounceTime    : TIME;
    CycleTime       : TIME;
END_VAR

VAR_OUTPUT
    VFD_RUN         : BOOL;
    PUMP_MAINT_DUE  : BOOL;
    PUMP_RUNTIME_ACC: LTIME;
END_VAR

VAR
    ViscosityDebounce : TON;
    tmpViscosityValid : BOOL;
END_VAR

// Single TON call per scan with correct input determined by E-stop
IF NOT PASTE_E_STOP_NC THEN
    ViscosityDebounce(IN := FALSE, PT := DebounceTime);
ELSE
    ViscosityDebounce(IN := VISCOSITY_OK, PT := DebounceTime);
END_IF;

tmpViscosityValid := ViscosityDebounce.Q;

IF NOT PASTE_E_STOP_NC THEN
    VFD_RUN := FALSE;
ELSE
    VFD_RUN := tmpViscosityValid;
END_IF;

IF VFD_RUN THEN
    PUMP_RUNTIME_ACC := PUMP_RUNTIME_ACC + TO_LTIME(CycleTime);
END_IF;

IF PUMP_RUNTIME_ACC >= T#500h THEN
    PUMP_MAINT_DUE := TRUE;
END_IF;

END_FUNCTION_BLOCK

(* ---- public-hard-03.candidate_01.st ---- *)
FUNCTION_BLOCK FB_RecipeManagement
VAR_INPUT
    addRecipe    : BOOL;
    deleteRecipe : BOOL;
    modifyRecipe : BOOL;
    queryRecipe  : BOOL;
    recipeIn     : ST_Recipe;
END_VAR

VAR_OUTPUT
    recipeAdded       : BOOL;
    recipeDeleted     : BOOL;
    recipeModified    : BOOL;
    recipeQueryResult : ST_Recipe;
    error             : BOOL;
    status            : WORD;
END_VAR

VAR_IN_OUT
    recipe : ARRAY[1..10] OF ST_Recipe;
END_VAR

VAR
    tmp_idx       : INT;
    tmp_foundIdx  : INT;
    tmp_emptyIdx  : INT;
END_VAR

// ENGINEERING_CONTRACT
(*
PUB001: Recipe management for production line control center
PUB002-006: CRUD operations on recipe database
PUB008: Array[1..10], recipeID=0 denotes empty slot, no duplicate IDs
PUB009: Query - not found => error=16#8001
PUB010: Add - duplicate => 16#8002, no slot => 16#8003
PUB011: Delete - not found => 16#8004
PUB012: Modify - not found => 16#8005
Output activation: recipeAdded/recipeDeleted/recipeModified = single-scan TRUE on success
Output retention: error/status persist until next operation; no latch
Same-scan priority: none required; sequential execution order preserved
*)

// CONTRACT_RULES
(* [] *)

recipeAdded := FALSE;
recipeDeleted := FALSE;
recipeModified := FALSE;
error := FALSE;
status := 16#0000;

tmp_foundIdx := 0;
tmp_emptyIdx := 0;

FOR tmp_idx := 1 TO 10 DO
    IF recipe[tmp_idx].recipeID = recipeIn.recipeID THEN
        tmp_foundIdx := tmp_idx;
    END_IF;
    IF recipe[tmp_idx].recipeID = 0 AND tmp_emptyIdx = 0 THEN
        tmp_emptyIdx := tmp_idx;
    END_IF;
END_FOR;

IF queryRecipe THEN
    IF tmp_foundIdx = 0 THEN
        error := TRUE;
        status := 16#8001;
    ELSE
        recipeQueryResult := recipe[tmp_foundIdx];
    END_IF;
ELSIF addRecipe THEN
    IF tmp_foundIdx <> 0 THEN
        error := TRUE;
        status := 16#8002;
    ELSIF tmp_emptyIdx = 0 THEN
        error := TRUE;
        status := 16#8003;
    ELSE
        recipe[tmp_emptyIdx] := recipeIn;
        recipeAdded := TRUE;
    END_IF;
ELSIF deleteRecipe THEN
    IF tmp_foundIdx = 0 THEN
        error := TRUE;
        status := 16#8004;
    ELSE
        recipe[tmp_foundIdx].recipeID := 0;
        recipeDeleted := TRUE;
    END_IF;
ELSIF modifyRecipe THEN
    IF tmp_foundIdx = 0 THEN
        error := TRUE;
        status := 16#8005;
    ELSE
        recipe[tmp_foundIdx] := recipeIn;
        recipeModified := TRUE;
    END_IF;
END_IF;

END_FUNCTION_BLOCK

(* ---- public-hard-03.candidate_02.st ---- *)
TYPE ST_Recipe :
STRUCT
    recipeID             : INT;
    ingredientType       : INT;
    ingredientRatio      : REAL;
    productionTemperature: REAL;
END_STRUCT
END_TYPE;

FUNCTION_BLOCK FB_RecipeManagement
VAR_INPUT
    addRecipe    : BOOL;
    deleteRecipe : BOOL;
    modifyRecipe : BOOL;
    queryRecipe  : BOOL;
    recipeIn     : ST_Recipe;
END_VAR

VAR_OUTPUT
    recipeAdded       : BOOL;
    recipeDeleted     : BOOL;
    recipeModified    : BOOL;
    recipeQueryResult : ST_Recipe;
    error             : BOOL;
    status            : WORD;
END_VAR

VAR_IN_OUT
    recipe : ARRAY[1..10] OF ST_Recipe;
END_VAR

VAR
    tmp_idx       : INT;
    tmp_foundIdx  : INT;
    tmp_emptyIdx  : INT;
END_VAR

// ENGINEERING_CONTRACT
(*
PUB001: Recipe management for production line control center
PUB002-006: CRUD operations on recipe database
PUB008: Array[1..10], recipeID=0 denotes empty slot, no duplicate IDs
PUB009: Query - not found => error=16#8001
PUB010: Add - duplicate => 16#8002, no slot => 16#8003
PUB011: Delete - not found => 16#8004
PUB012: Modify - not found => 16#8005
Output activation: recipeAdded/recipeDeleted/recipeModified = single-scan TRUE on success
Output retention: error/status persist until next operation; no latch
Same-scan priority: none required; sequential execution order preserved
*)

// CONTRACT_RULES
(* [] *)

recipeAdded := FALSE;
recipeDeleted := FALSE;
recipeModified := FALSE;
error := FALSE;
status := 16#0000;

tmp_foundIdx := 0;
tmp_emptyIdx := 0;

FOR tmp_idx := 1 TO 10 DO
    IF recipe[tmp_idx].recipeID = recipeIn.recipeID THEN
        tmp_foundIdx := tmp_idx;
    END_IF;
    IF recipe[tmp_idx].recipeID = 0 AND tmp_emptyIdx = 0 THEN
        tmp_emptyIdx := tmp_idx;
    END_IF;
END_FOR;

IF queryRecipe THEN
    IF tmp_foundIdx = 0 THEN
        error := TRUE;
        status := 16#8001;
    ELSE
        recipeQueryResult := recipe[tmp_foundIdx];
    END_IF;
ELSIF addRecipe THEN
    IF tmp_foundIdx <> 0 THEN
        error := TRUE;
        status := 16#8002;
    ELSIF tmp_emptyIdx = 0 THEN
        error := TRUE;
        status := 16#8003;
    ELSE
        recipe[tmp_emptyIdx] := recipeIn;
        recipeAdded := TRUE;
    END_IF;
ELSIF deleteRecipe THEN
    IF tmp_foundIdx = 0 THEN
        error := TRUE;
        status := 16#8004;
    ELSE
        recipe[tmp_foundIdx].recipeID := 0;
        recipeDeleted := TRUE;
    END_IF;
ELSIF modifyRecipe THEN
    IF tmp_foundIdx = 0 THEN
        error := TRUE;
        status := 16#8005;
    ELSE
        recipe[tmp_foundIdx] := recipeIn;
        recipeModified := TRUE;
    END_IF;
END_IF;

END_FUNCTION_BLOCK

(* ---- public-hard-03.candidate_03.st ---- *)
TYPE ST_Recipe :
STRUCT
    recipeID             : INT;
    ingredientType       : INT;
    ingredientRatio      : REAL;
    productionTemperature: REAL;
END_STRUCT
END_TYPE;

FUNCTION_BLOCK FB_RecipeManagement
VAR_INPUT
    addRecipe    : BOOL;
    deleteRecipe : BOOL;
    modifyRecipe : BOOL;
    queryRecipe  : BOOL;
    recipeIn     : ST_Recipe;
END_VAR

VAR_OUTPUT
    recipeAdded       : BOOL;
    recipeDeleted     : BOOL;
    recipeModified    : BOOL;
    recipeQueryResult : ST_Recipe;
    error             : BOOL;
    status            : WORD;
END_VAR

VAR_IN_OUT
    recipe : ARRAY[1..10] OF ST_Recipe;
END_VAR

VAR
    tmp_idx       : INT;
    tmp_foundIdx  : INT;
    tmp_emptyIdx  : INT;
END_VAR

// ENGINEERING_CONTRACT
(*
PUB001: Recipe management for production line control center
PUB002-006: CRUD operations on recipe database
PUB008: Array[1..10], recipeID=0 denotes empty slot, no duplicate IDs
PUB009: Query - not found => error=TRUE, status=16#8001
PUB010: Add - duplicate => 16#8002, no slot => 16#8003, else store at smallest empty index
PUB011: Delete - not found => 16#8004, else set recipeID=0
PUB012: Modify - not found => 16#8005, else replace entire recipe
Output activation: recipeAdded/recipeDeleted/recipeModified = single-scan TRUE on success
Output retention: error/status persist until next operation; no persistent latch
Same-scan priority: IF/ELSIF chain order = queryRecipe > addRecipe > deleteRecipe > modifyRecipe
Units/boundaries: recipe array[1..10], recipeID=INT (0=empty), ratio/temp=REAL
*)

// CONTRACT_RULES
(* [] *)

recipeAdded := FALSE;
recipeDeleted := FALSE;
recipeModified := FALSE;
error := FALSE;
status := 16#0000;

tmp_foundIdx := 0;
tmp_emptyIdx := 0;

FOR tmp_idx := 1 TO 10 DO
    IF recipe[tmp_idx].recipeID = recipeIn.recipeID THEN
        tmp_foundIdx := tmp_idx;
    END_IF;
    IF recipe[tmp_idx].recipeID = 0 AND tmp_emptyIdx = 0 THEN
        tmp_emptyIdx := tmp_idx;
    END_IF;
END_FOR;

IF queryRecipe THEN
    IF tmp_foundIdx = 0 THEN
        error := TRUE;
        status := 16#8001;
    ELSE
        recipeQueryResult := recipe[tmp_foundIdx];
    END_IF;
ELSIF addRecipe THEN
    IF tmp_foundIdx <> 0 THEN
        error := TRUE;
        status := 16#8002;
    ELSIF tmp_emptyIdx = 0 THEN
        error := TRUE;
        status := 16#8003;
    ELSE
        recipe[tmp_emptyIdx] := recipeIn;
        recipeAdded := TRUE;
    END_IF;
ELSIF deleteRecipe THEN
    IF tmp_foundIdx = 0 THEN
        error := TRUE;
        status := 16#8004;
    ELSE
        recipe[tmp_foundIdx].recipeID := 0;
        recipeDeleted := TRUE;
    END_IF;
ELSIF modifyRecipe THEN
    IF tmp_foundIdx = 0 THEN
        error := TRUE;
        status := 16#8005;
    ELSE
        recipe[tmp_foundIdx] := recipeIn;
        recipeModified := TRUE;
    END_IF;
END_IF;

END_FUNCTION_BLOCK

(* ---- public-hard-03.candidate_04.st ---- *)
TYPE ST_Recipe :
STRUCT
    recipeID             : INT;
    ingredientType       : INT;
    ingredientRatio      : REAL;
    productionTemperature: REAL;
END_STRUCT
END_TYPE;

FUNCTION_BLOCK FB_RecipeManagement
VAR_INPUT
    addRecipe    : BOOL;
    deleteRecipe : BOOL;
    modifyRecipe : BOOL;
    queryRecipe  : BOOL;
    recipeIn     : ST_Recipe;
END_VAR

VAR_OUTPUT
    recipeAdded       : BOOL;
    recipeDeleted     : BOOL;
    recipeModified    : BOOL;
    recipeQueryResult : ST_Recipe;
    error             : BOOL;
    status            : WORD;
END_VAR

VAR_IN_OUT
    recipe : ARRAY[1..10] OF ST_Recipe;
END_VAR

VAR
    tmp_idx       : INT;
    tmp_foundIdx  : INT;
    tmp_emptyIdx  : INT;
END_VAR

// ENGINEERING_CONTRACT
(*
PUB001: Recipe management for production line control center
PUB002-006: CRUD operations on recipe database
PUB008: Array[1..10], recipeID=0 denotes empty slot, no duplicate IDs
PUB009: Query - not found => error=16#8001
PUB010: Add - duplicate => 16#8002, no slot => 16#8003
PUB011: Delete - not found => 16#8004
PUB012: Modify - not found => 16#8005
Output activation: recipeAdded/recipeDeleted/recipeModified = single-scan TRUE on success
Output retention: error/status persist until next operation; no latch
Same-scan priority: ELSIF order defines precedence (query > add > delete > modify)
*)

// CONTRACT_RULES
(* [] *)

recipeAdded   := FALSE;
recipeDeleted := FALSE;
recipeModified := FALSE;
error         := FALSE;
status        := 16#0000;

tmp_foundIdx := 0;
tmp_emptyIdx := 0;

FOR tmp_idx := 1 TO 10 DO
    IF recipe[tmp_idx].recipeID = recipeIn.recipeID THEN
        tmp_foundIdx := tmp_idx;
    END_IF;
    IF recipe[tmp_idx].recipeID = 0 AND tmp_emptyIdx = 0 THEN
        tmp_emptyIdx := tmp_idx;
    END_IF;
END_FOR;

IF queryRecipe THEN
    IF tmp_foundIdx = 0 THEN
        error := TRUE;
        status := 16#8001;
    ELSE
        recipeQueryResult := recipe[tmp_foundIdx];
    END_IF;
ELSIF addRecipe THEN
    IF tmp_foundIdx <> 0 THEN
        error := TRUE;
        status := 16#8002;
    ELSIF tmp_emptyIdx = 0 THEN
        error := TRUE;
        status := 16#8003;
    ELSE
        recipe[tmp_emptyIdx] := recipeIn;
        recipeAdded := TRUE;
    END_IF;
ELSIF deleteRecipe THEN
    IF tmp_foundIdx = 0 THEN
        error := TRUE;
        status := 16#8004;
    ELSE
        recipe[tmp_foundIdx].recipeID := 0;
        recipeDeleted := TRUE;
    END_IF;
ELSIF modifyRecipe THEN
    IF tmp_foundIdx = 0 THEN
        error := TRUE;
        status := 16#8005;
    ELSE
        recipe[tmp_foundIdx] := recipeIn;
        recipeModified := TRUE;
    END_IF;
END_IF;

END_FUNCTION_BLOCK

(* ---- public-hard-03.raw_candidate_01.st ---- *)
FUNCTION_BLOCK FB_RecipeManagement
VAR_INPUT
    addRecipe    : BOOL;
    deleteRecipe : BOOL;
    modifyRecipe : BOOL;
    queryRecipe  : BOOL;
    recipeIn     : ST_Recipe;
END_VAR

VAR_OUTPUT
    recipeAdded       : BOOL;
    recipeDeleted     : BOOL;
    recipeModified    : BOOL;
    recipeQueryResult : ST_Recipe;
    error             : BOOL;
    status            : WORD;
END_VAR

VAR_IN_OUT
    recipe : ARRAY[1..10] OF ST_Recipe;
END_VAR

VAR
    tmp_idx       : INT;
    tmp_foundIdx  : INT;
    tmp_emptyIdx  : INT;
END_VAR

// ENGINEERING_CONTRACT
(*
PUB001: Recipe management for production line control center
PUB002-006: CRUD operations on recipe database
PUB008: Array[1..10], recipeID=0 denotes empty slot, no duplicate IDs
PUB009: Query - not found => error=16#8001
PUB010: Add - duplicate => 16#8002, no slot => 16#8003
PUB011: Delete - not found => 16#8004
PUB012: Modify - not found => 16#8005
Output activation: recipeAdded/recipeDeleted/recipeModified = single-scan TRUE on success
Output retention: error/status persist until next operation; no latch
Same-scan priority: none required; sequential execution order preserved
*)

// CONTRACT_RULES
(* [] *)

recipeAdded := FALSE;
recipeDeleted := FALSE;
recipeModified := FALSE;
error := FALSE;
status := 16#0000;

tmp_foundIdx := 0;
tmp_emptyIdx := 0;

FOR tmp_idx := 1 TO 10 DO
    IF recipe[tmp_idx].recipeID = recipeIn.recipeID THEN
        tmp_foundIdx := tmp_idx;
    END_IF
    IF recipe[tmp_idx].recipeID = 0 AND tmp_emptyIdx = 0 THEN
        tmp_emptyIdx := tmp_idx;
    END_IF
END_FOR

IF queryRecipe THEN
    IF tmp_foundIdx = 0 THEN
        error := TRUE;
        status := 16#8001;
    ELSE
        recipeQueryResult := recipe[tmp_foundIdx];
    END_IF;
ELSIF addRecipe THEN
    IF tmp_foundIdx <> 0 THEN
        error := TRUE;
        status := 16#8002;
    ELSIF tmp_emptyIdx = 0 THEN
        error := TRUE;
        status := 16#8003;
    ELSE
        recipe[tmp_emptyIdx] := recipeIn;
        recipeAdded := TRUE;
    END_IF;
ELSIF deleteRecipe THEN
    IF tmp_foundIdx = 0 THEN
        error := TRUE;
        status := 16#8004;
    ELSE
        recipe[tmp_foundIdx].recipeID := 0;
        recipeDeleted := TRUE;
    END_IF;
ELSIF modifyRecipe THEN
    IF tmp_foundIdx = 0 THEN
        error := TRUE;
        status := 16#8005;
    ELSE
        recipe[tmp_foundIdx] := recipeIn;
        recipeModified := TRUE;
    END_IF;
END_IF;

END_FUNCTION_BLOCK

(* ---- public-hard-03.raw_candidate_02.st ---- *)
TYPE ST_Recipe :
STRUCT
    recipeID             : INT;
    ingredientType       : INT;
    ingredientRatio      : REAL;
    productionTemperature: REAL;
END_STRUCT
END_TYPE

FUNCTION_BLOCK FB_RecipeManagement
VAR_INPUT
    addRecipe    : BOOL;
    deleteRecipe : BOOL;
    modifyRecipe : BOOL;
    queryRecipe  : BOOL;
    recipeIn     : ST_Recipe;
END_VAR

VAR_OUTPUT
    recipeAdded       : BOOL;
    recipeDeleted     : BOOL;
    recipeModified    : BOOL;
    recipeQueryResult : ST_Recipe;
    error             : BOOL;
    status            : WORD;
END_VAR

VAR_IN_OUT
    recipe : ARRAY[1..10] OF ST_Recipe;
END_VAR

VAR
    tmp_idx       : INT;
    tmp_foundIdx  : INT;
    tmp_emptyIdx  : INT;
END_VAR

// ENGINEERING_CONTRACT
(*
PUB001: Recipe management for production line control center
PUB002-006: CRUD operations on recipe database
PUB008: Array[1..10], recipeID=0 denotes empty slot, no duplicate IDs
PUB009: Query - not found => error=16#8001
PUB010: Add - duplicate => 16#8002, no slot => 16#8003
PUB011: Delete - not found => 16#8004
PUB012: Modify - not found => 16#8005
Output activation: recipeAdded/recipeDeleted/recipeModified = single-scan TRUE on success
Output retention: error/status persist until next operation; no latch
Same-scan priority: none required; sequential execution order preserved
*)

// CONTRACT_RULES
(* [] *)

recipeAdded := FALSE;
recipeDeleted := FALSE;
recipeModified := FALSE;
error := FALSE;
status := 16#0000;

tmp_foundIdx := 0;
tmp_emptyIdx := 0;

FOR tmp_idx := 1 TO 10 DO
    IF recipe[tmp_idx].recipeID = recipeIn.recipeID THEN
        tmp_foundIdx := tmp_idx;
    END_IF;
    IF recipe[tmp_idx].recipeID = 0 AND tmp_emptyIdx = 0 THEN
        tmp_emptyIdx := tmp_idx;
    END_IF;
END_FOR;

IF queryRecipe THEN
    IF tmp_foundIdx = 0 THEN
        error := TRUE;
        status := 16#8001;
    ELSE
        recipeQueryResult := recipe[tmp_foundIdx];
    END_IF;
ELSIF addRecipe THEN
    IF tmp_foundIdx <> 0 THEN
        error := TRUE;
        status := 16#8002;
    ELSIF tmp_emptyIdx = 0 THEN
        error := TRUE;
        status := 16#8003;
    ELSE
        recipe[tmp_emptyIdx] := recipeIn;
        recipeAdded := TRUE;
    END_IF;
ELSIF deleteRecipe THEN
    IF tmp_foundIdx = 0 THEN
        error := TRUE;
        status := 16#8004;
    ELSE
        recipe[tmp_foundIdx].recipeID := 0;
        recipeDeleted := TRUE;
    END_IF;
ELSIF modifyRecipe THEN
    IF tmp_foundIdx = 0 THEN
        error := TRUE;
        status := 16#8005;
    ELSE
        recipe[tmp_foundIdx] := recipeIn;
        recipeModified := TRUE;
    END_IF;
END_IF;

END_FUNCTION_BLOCK

(* ---- public-hard-03.raw_candidate_03.st ---- *)
TYPE ST_Recipe :
STRUCT
    recipeID             : INT;
    ingredientType       : INT;
    ingredientRatio      : REAL;
    productionTemperature: REAL;
END_STRUCT
END_TYPE

FUNCTION_BLOCK FB_RecipeManagement
VAR_INPUT
    addRecipe    : BOOL;
    deleteRecipe : BOOL;
    modifyRecipe : BOOL;
    queryRecipe  : BOOL;
    recipeIn     : ST_Recipe;
END_VAR

VAR_OUTPUT
    recipeAdded       : BOOL;
    recipeDeleted     : BOOL;
    recipeModified    : BOOL;
    recipeQueryResult : ST_Recipe;
    error             : BOOL;
    status            : WORD;
END_VAR

VAR_IN_OUT
    recipe : ARRAY[1..10] OF ST_Recipe;
END_VAR

VAR
    tmp_idx       : INT;
    tmp_foundIdx  : INT;
    tmp_emptyIdx  : INT;
END_VAR

// ENGINEERING_CONTRACT
(*
PUB001: Recipe management for production line control center
PUB002-006: CRUD operations on recipe database
PUB008: Array[1..10], recipeID=0 denotes empty slot, no duplicate IDs
PUB009: Query - not found => error=TRUE, status=16#8001
PUB010: Add - duplicate => 16#8002, no slot => 16#8003, else store at smallest empty index
PUB011: Delete - not found => 16#8004, else set recipeID=0
PUB012: Modify - not found => 16#8005, else replace entire recipe
Output activation: recipeAdded/recipeDeleted/recipeModified = single-scan TRUE on success
Output retention: error/status persist until next operation; no persistent latch
Same-scan priority: IF/ELSIF chain order = queryRecipe > addRecipe > deleteRecipe > modifyRecipe
Units/boundaries: recipe array[1..10], recipeID=INT (0=empty), ratio/temp=REAL
*)

// CONTRACT_RULES
(* [] *)

recipeAdded := FALSE;
recipeDeleted := FALSE;
recipeModified := FALSE;
error := FALSE;
status := 16#0000;

tmp_foundIdx := 0;
tmp_emptyIdx := 0;

FOR tmp_idx := 1 TO 10 DO
    IF recipe[tmp_idx].recipeID = recipeIn.recipeID THEN
        tmp_foundIdx := tmp_idx;
    END_IF;
    IF recipe[tmp_idx].recipeID = 0 AND tmp_emptyIdx = 0 THEN
        tmp_emptyIdx := tmp_idx;
    END_IF;
END_FOR;

IF queryRecipe THEN
    IF tmp_foundIdx = 0 THEN
        error := TRUE;
        status := 16#8001;
    ELSE
        recipeQueryResult := recipe[tmp_foundIdx];
    END_IF;
ELSIF addRecipe THEN
    IF tmp_foundIdx <> 0 THEN
        error := TRUE;
        status := 16#8002;
    ELSIF tmp_emptyIdx = 0 THEN
        error := TRUE;
        status := 16#8003;
    ELSE
        recipe[tmp_emptyIdx] := recipeIn;
        recipeAdded := TRUE;
    END_IF;
ELSIF deleteRecipe THEN
    IF tmp_foundIdx = 0 THEN
        error := TRUE;
        status := 16#8004;
    ELSE
        recipe[tmp_foundIdx].recipeID := 0;
        recipeDeleted := TRUE;
    END_IF;
ELSIF modifyRecipe THEN
    IF tmp_foundIdx = 0 THEN
        error := TRUE;
        status := 16#8005;
    ELSE
        recipe[tmp_foundIdx] := recipeIn;
        recipeModified := TRUE;
    END_IF;
END_IF;

END_FUNCTION_BLOCK

(* ---- public-hard-03.raw_candidate_04.st ---- *)
TYPE ST_Recipe :
STRUCT
    recipeID             : INT;
    ingredientType       : INT;
    ingredientRatio      : REAL;
    productionTemperature: REAL;
END_STRUCT
END_TYPE

FUNCTION_BLOCK FB_RecipeManagement
VAR_INPUT
    addRecipe    : BOOL;
    deleteRecipe : BOOL;
    modifyRecipe : BOOL;
    queryRecipe  : BOOL;
    recipeIn     : ST_Recipe;
END_VAR

VAR_OUTPUT
    recipeAdded       : BOOL;
    recipeDeleted     : BOOL;
    recipeModified    : BOOL;
    recipeQueryResult : ST_Recipe;
    error             : BOOL;
    status            : WORD;
END_VAR

VAR_IN_OUT
    recipe : ARRAY[1..10] OF ST_Recipe;
END_VAR

VAR
    tmp_idx       : INT;
    tmp_foundIdx  : INT;
    tmp_emptyIdx  : INT;
END_VAR

// ENGINEERING_CONTRACT
(*
PUB001: Recipe management for production line control center
PUB002-006: CRUD operations on recipe database
PUB008: Array[1..10], recipeID=0 denotes empty slot, no duplicate IDs
PUB009: Query - not found => error=16#8001
PUB010: Add - duplicate => 16#8002, no slot => 16#8003
PUB011: Delete - not found => 16#8004
PUB012: Modify - not found => 16#8005
Output activation: recipeAdded/recipeDeleted/recipeModified = single-scan TRUE on success
Output retention: error/status persist until next operation; no latch
Same-scan priority: ELSIF order defines precedence (query > add > delete > modify)
*)

// CONTRACT_RULES
(* [] *)

recipeAdded   := FALSE;
recipeDeleted := FALSE;
recipeModified := FALSE;
error         := FALSE;
status        := 16#0000;

tmp_foundIdx := 0;
tmp_emptyIdx := 0;

FOR tmp_idx := 1 TO 10 DO
    IF recipe[tmp_idx].recipeID = recipeIn.recipeID THEN
        tmp_foundIdx := tmp_idx;
    END_IF;
    IF recipe[tmp_idx].recipeID = 0 AND tmp_emptyIdx = 0 THEN
        tmp_emptyIdx := tmp_idx;
    END_IF;
END_FOR;

IF queryRecipe THEN
    IF tmp_foundIdx = 0 THEN
        error := TRUE;
        status := 16#8001;
    ELSE
        recipeQueryResult := recipe[tmp_foundIdx];
    END_IF;
ELSIF addRecipe THEN
    IF tmp_foundIdx <> 0 THEN
        error := TRUE;
        status := 16#8002;
    ELSIF tmp_emptyIdx = 0 THEN
        error := TRUE;
        status := 16#8003;
    ELSE
        recipe[tmp_emptyIdx] := recipeIn;
        recipeAdded := TRUE;
    END_IF;
ELSIF deleteRecipe THEN
    IF tmp_foundIdx = 0 THEN
        error := TRUE;
        status := 16#8004;
    ELSE
        recipe[tmp_foundIdx].recipeID := 0;
        recipeDeleted := TRUE;
    END_IF;
ELSIF modifyRecipe THEN
    IF tmp_foundIdx = 0 THEN
        error := TRUE;
        status := 16#8005;
    ELSE
        recipe[tmp_foundIdx] := recipeIn;
        recipeModified := TRUE;
    END_IF;
END_IF;

END_FUNCTION_BLOCK

(* ---- public-medium-03.candidate_01.st ---- *)
{engineer}
(* CONTRACT_RULES [] *)
(* ENGINEERING_CONTRACT
 * ID              | Activation                    | Retention         | Reset/Deactivation | Priority   | Units/Boundaries
 * ----------------------------------------------------------------------------------------------------------------------------------
 * average         | cyclicExecution=TRUE          | Until next value  | reset=TRUE         | Same-scan  | LREAL, output
 *                 | trigger rising edge           |                   |                    |            |
 * windowSizeReached | currentWindowSize=windowSize | Until reset       | reset=TRUE         | Same-scan  | BOOL, output
 * error           | windowSize < 1 OR > 100       | Until reset       | reset=TRUE         | Same-scan  | BOOL, output
 * status          | Derived from windowSize check | Until reset       | reset=TRUE         | Same-scan  | WORD: 16#0000 or 16#8200
 *
 * Data buffer: circular buffer of 100 LREAL entries (max window size)
 * Sum maintained incrementally for O(1) average calculation
 * PUB001, PUB002, PUB003, PUB004, PUB006, PUB007
 *)
FUNCTION_BLOCK FB_MovingAverage
VAR_INPUT
    cyclicExecution : BOOL;
    trigger : BOOL;
    value : LREAL;
    windowSize : INT;
    reset : BOOL;
END_VAR
VAR_OUTPUT
    average : LREAL := 0.0;
    windowSizeReached : BOOL := FALSE;
    error : BOOL := FALSE;
    status : WORD := 16#0000;
END_VAR
VAR
    dataBuffer : ARRAY[1..100] OF LREAL;
    bufferIndex : INT := 0;
    currentWindowSize : INT := 0;
    sum : LREAL := 0.0;
    lastTrigger : BOOL := FALSE;
END_VAR

// Reset handling
IF reset THEN
    bufferIndex := 0;
    currentWindowSize := 0;
    sum := 0.0;
    average := 0.0;
    windowSizeReached := FALSE;
    error := FALSE;
    status := 16#0000;
    lastTrigger := FALSE;
    RETURN;
END_IF;

// Validate window size
IF windowSize < 1 OR windowSize > 100 THEN
    error := TRUE;
    status := 16#8200;
    RETURN;
END_IF;

// Cyclic execution takes priority over trigger
IF cyclicExecution THEN
    IF currentWindowSize >= windowSize THEN
        // Window is full, replace oldest value
        bufferIndex := (bufferIndex MOD windowSize) + 1;
        sum := sum - dataBuffer[bufferIndex] + value;
        average := sum / TO_LREAL(windowSize);
    ELSE
        // Window not yet full, add new value
        bufferIndex := bufferIndex + 1;
        dataBuffer[bufferIndex] := value;
        sum := sum + value;
        currentWindowSize := bufferIndex;
        average := sum / TO_LREAL(currentWindowSize);
    END_IF;

    windowSizeReached := (currentWindowSize >= windowSize);
    error := FALSE;
    status := 16#0000;
    RETURN;
END_IF;

// Trigger-based execution on rising edge
IF trigger AND NOT lastTrigger THEN
    IF currentWindowSize >= windowSize THEN
        // Window is full, replace oldest value
        bufferIndex := (bufferIndex MOD windowSize) + 1;
        sum := sum - dataBuffer[bufferIndex] + value;
        average := sum / TO_LREAL(windowSize);
    ELSE
        // Window not yet full, add new value
        bufferIndex := bufferIndex + 1;
        dataBuffer[bufferIndex] := value;
        sum := sum + value;
        currentWindowSize := bufferIndex;
        average := sum / TO_LREAL(currentWindowSize);
    END_IF;

    windowSizeReached := (currentWindowSize >= windowSize);
    error := FALSE;
    status := 16#0000;
END_IF;

lastTrigger := trigger;
END_FUNCTION_BLOCK

(* ---- public-medium-03.raw_candidate_01.st ---- *)
{engineer}
(* CONTRACT_RULES [] *)
(* ENGINEERING_CONTRACT
 * ID              | Activation                    | Retention         | Reset/Deactivation | Priority   | Units/Boundaries
 * ----------------------------------------------------------------------------------------------------------------------------------
 * average         | cyclicExecution=TRUE          | Until next value  | reset=TRUE         | Same-scan  | LREAL, output
 *                 | trigger rising edge           |                   |                    |            |
 * windowSizeReached | currentWindowSize=windowSize | Until reset       | reset=TRUE         | Same-scan  | BOOL, output
 * error           | windowSize < 1 OR > 100       | Until reset       | reset=TRUE         | Same-scan  | BOOL, output
 * status          | Derived from windowSize check | Until reset       | reset=TRUE         | Same-scan  | WORD: 16#0000 or 16#8200
 *
 * Data buffer: circular buffer of 100 LREAL entries (max window size)
 * Sum maintained incrementally for O(1) average calculation
 * PUB001, PUB002, PUB003, PUB004, PUB006, PUB007
 *)
FUNCTION_BLOCK FB_MovingAverage
VAR_INPUT
    cyclicExecution : BOOL;
    trigger : BOOL;
    value : LREAL;
    windowSize : INT;
    reset : BOOL;
END_VAR
VAR_OUTPUT
    average : LREAL := 0.0;
    windowSizeReached : BOOL := FALSE;
    error : BOOL := FALSE;
    status : WORD := 16#0000;
END_VAR
VAR
    dataBuffer : ARRAY[1..100] OF LREAL;
    bufferIndex : INT := 0;
    currentWindowSize : INT := 0;
    sum : LREAL := 0.0;
    lastTrigger : BOOL := FALSE;
END_VAR

// Reset handling
IF reset THEN
    bufferIndex := 0;
    currentWindowSize := 0;
    sum := 0.0;
    average := 0.0;
    windowSizeReached := FALSE;
    error := FALSE;
    status := 16#0000;
    lastTrigger := FALSE;
    RETURN;
END_IF;

// Validate window size
IF windowSize < 1 OR windowSize > 100 THEN
    error := TRUE;
    status := 16#8200;
    RETURN;
END_IF;

// Cyclic execution takes priority over trigger
IF cyclicExecution THEN
    IF currentWindowSize >= windowSize THEN
        // Window is full, replace oldest value
        bufferIndex := (bufferIndex MOD windowSize) + 1;
        sum := sum - dataBuffer[bufferIndex] + value;
        average := sum / TO_LREAL(windowSize);
    ELSE
        // Window not yet full, add new value
        bufferIndex := bufferIndex + 1;
        dataBuffer[bufferIndex] := value;
        sum := sum + value;
        currentWindowSize := bufferIndex;
        average := sum / TO_LREAL(currentWindowSize);
    END_IF;

    windowSizeReached := (currentWindowSize >= windowSize);
    error := FALSE;
    status := 16#0000;
    RETURN;
END_IF;

// Trigger-based execution on rising edge
IF trigger AND NOT lastTrigger THEN
    IF currentWindowSize >= windowSize THEN
        // Window is full, replace oldest value
        bufferIndex := (bufferIndex MOD windowSize) + 1;
        sum := sum - dataBuffer[bufferIndex] + value;
        average := sum / TO_LREAL(windowSize);
    ELSE
        // Window not yet full, add new value
        bufferIndex := bufferIndex + 1;
        dataBuffer[bufferIndex] := value;
        sum := sum + value;
        currentWindowSize := bufferIndex;
        average := sum / TO_LREAL(currentWindowSize);
    END_IF;

    windowSizeReached := (currentWindowSize >= windowSize);
    error := FALSE;
    status := 16#0000;
END_IF;

lastTrigger := trigger;
END_FUNCTION_BLOCK

(* ---- public-medium-04.candidate_01.st ---- *)
FUNCTION_BLOCK FB_TemperatureControl
VAR_INPUT
    TemperatureSensorInput : REAL;
    SetTemperature : REAL;
END_VAR
VAR_OUTPUT
    CurrentTemperature : REAL;
    SetTempDisplay : REAL;
    HeaterStatus : BOOL;
    OverheatProtection : BOOL;
    HeaterOutput : BOOL;
END_VAR
VAR
    HeaterOnRequest : BOOL;
    OverheatTimer : TON;
    OverheatCooldownTimer : TON;
    tmp_SensorFault : BOOL;
    tmp_HeaterShouldBeOn : BOOL;
END_VAR

(* ENGINEERING_CONTRACT
 * ============================================================
 * Outputs & State Groups:
 * -----------------------------------------------------------
 * HeaterOutput (BOOL, output):
 *   - Activation: Set TRUE when temp < set, no fault, no overheat
 *   - Retention: Maintained TRUE across scans while conditions hold
 *   - Explicit Reset: Set FALSE by fault detection OR overheat trigger
 *   - Same-scan Priority: Fault > Overheat > Temperature comparison
 *   - Units: Boolean on/off signal
 * -----------------------------------------------------------
 * OverheatProtection (BOOL, output):
 *   - Activation: Set TRUE after heater runs continuously > 5s (PUB006)
 *   - Retention: Held TRUE for mandatory 3s cooldown period (PUB006)
 *   - Explicit Reset: Cleared automatically after 3s elapses
 *   - Same-scan Priority: Timer expiry drives reset after 3s
 *   - Units: Boolean flag (TRUE = protection latched)
 * -----------------------------------------------------------
 * CurrentTemperature / SetTempDisplay (REAL, output):
 *   - Activation: Assigned every scan from inputs
 *   - Retention: No retention; mirrors inputs each scan
 *   - Explicit Reset: N/A (always reflects current values)
 *   - Same-scan Priority: Direct assignment
 *   - Units: degrees (temperature values, PUB002/PUB007)
 * -----------------------------------------------------------
 * HeaterStatus (BOOL, output):
 *   - Activation: Mirrors HeaterOutput value each scan
 *   - Retention: Reflects current heater state
 *   - Explicit Reset: Same as HeaterOutput
 *   - Units: Boolean status indicator (PUB007)
 * ============================================================
 * CONTRACT_RULES []
 * ============================================================ *)

tmp_SensorFault := (TemperatureSensorInput < 0.0) OR (TemperatureSensorInput > 100.0);

CurrentTemperature := TemperatureSensorInput;
SetTempDisplay := SetTemperature;

IF tmp_SensorFault THEN
    HeaterOnRequest := FALSE;
ELSIF OverheatProtection THEN
    HeaterOnRequest := FALSE;
ELSE
    tmp_HeaterShouldBeOn := (TemperatureSensorInput < SetTemperature);
    HeaterOnRequest := tmp_HeaterShouldBeOn;
END_IF;

OverheatTimer(IN := HeaterOnRequest AND NOT OverheatProtection,
              PT := T#5S);

IF OverheatTimer.Q THEN
    OverheatProtection := TRUE;
END_IF;

OverheatCooldownTimer(IN := OverheatProtection,
                      PT := T#3S);

IF OverheatCooldownTimer.Q THEN
    OverheatProtection := FALSE;
END_IF;

HeaterOutput := HeaterOnRequest;
HeaterStatus := HeaterOutput;

END_FUNCTION_BLOCK

(* ---- public-medium-04.candidate_02.st ---- *)
FUNCTION_BLOCK FB_TemperatureControl
VAR_INPUT
    TemperatureSensorInput : REAL;
    SetTemperature : REAL;
END_VAR
VAR_OUTPUT
    CurrentTemperature : REAL;
    SetTempDisplay : REAL;
    HeaterStatus : BOOL;
    OverheatProtection : BOOL;
    HeaterOutput : BOOL;
END_VAR
VAR
    HeaterOnRequest : BOOL;
    OverheatTimer : TON;
    CooldownTimer : TON;
    tmp_SensorFault : BOOL;
    tmp_HeaterShouldBeOn : BOOL;
END_VAR

(* ENGINEERING_CONTRACT
 * ============================================================
 * Outputs & State Groups:
 * -----------------------------------------------------------
 * HeaterOutput (BOOL, output):
 *   - Activation: Set TRUE when temp < set, no fault, no overheat
 *   - Retention: Maintained TRUE across scans while conditions hold
 *   - Explicit Reset: Set FALSE by fault detection OR overheat trigger
 *   - Same-scan Priority: Fault > Overheat > Temperature comparison
 *   - Units: Boolean on/off signal
 * -----------------------------------------------------------
 * OverheatProtection (BOOL, output):
 *   - Activation: Set TRUE after heater runs continuously > 5s (PUB006)
 *   - Retention: Held TRUE for mandatory 3s cooldown period (PUB006)
 *   - Explicit Reset: Cleared automatically after 3s elapses
 *   - Same-scan Priority: Timer expiry drives reset after 3s
 *   - Units: Boolean flag (TRUE = protection latched)
 * -----------------------------------------------------------
 * CurrentTemperature / SetTempDisplay (REAL, output):
 *   - Activation: Assigned every scan from inputs
 *   - Retention: No retention; mirrors inputs each scan
 *   - Explicit Reset: N/A (always reflects current values)
 *   - Units: degrees (temperature values, PUB002/PUB007)
 * -----------------------------------------------------------
 * HeaterStatus (BOOL, output):
 *   - Activation: Mirrors HeaterOutput value each scan
 *   - Retention: Reflects current heater state
 *   - Units: Boolean status indicator (PUB007)
 * ============================================================
 * CONTRACT_RULES []
 * ============================================================ *)

tmp_SensorFault := (TemperatureSensorInput < 0.0) OR (TemperatureSensorInput > 100.0);

CurrentTemperature := TemperatureSensorInput;
SetTempDisplay := SetTemperature;

IF tmp_SensorFault THEN
    HeaterOnRequest := FALSE;
ELSIF OverheatProtection THEN
    HeaterOnRequest := FALSE;
ELSE
    tmp_HeaterShouldBeOn := (TemperatureSensorInput < SetTemperature);
    HeaterOnRequest := tmp_HeaterShouldBeOn;
END_IF;

OverheatTimer(IN := HeaterOnRequest AND NOT OverheatProtection,
              PT := T#5S);

IF OverheatTimer.Q THEN
    OverheatProtection := TRUE;
END_IF;

CooldownTimer(IN := OverheatProtection,
              PT := T#3S);

IF CooldownTimer.Q THEN
    OverheatProtection := FALSE;
END_IF;

HeaterOutput := HeaterOnRequest;
HeaterStatus := HeaterOutput;

END_FUNCTION_BLOCK

(* ---- public-medium-04.candidate_03.st ---- *)
FUNCTION_BLOCK FB_TemperatureControl
VAR_INPUT
    TemperatureSensorInput : REAL;
    SetTemperature : REAL;
END_VAR
VAR_OUTPUT
    CurrentTemperature : REAL;
    SetTempDisplay : REAL;
    HeaterStatus : BOOL;
    OverheatProtection : BOOL;
    HeaterOutput : BOOL;
END_VAR
VAR
    HeaterOnRequest : BOOL;
    OverheatTimer : TON;
    OverheatCooldownTimer : TON;
    tmp_SensorFault : BOOL;
END_VAR

(* ENGINEERING_CONTRACT
 * ============================================================
 * Outputs & State Groups:
 * -----------------------------------------------------------
 * HeaterOutput (BOOL, output):
 *   - Activation: Set TRUE when temp < set, no fault, no overheat
 *   - Retention: Maintained TRUE across scans while conditions hold
 *   - Explicit Reset: Set FALSE by fault OR overheat trigger (same-scan)
 *   - Same-scan Priority: OverheatProtection > Fault > Temperature
 *   - Units: Boolean on/off signal
 * -----------------------------------------------------------
 * OverheatProtection (BOOL, output):
 *   - Activation: Set TRUE after heater runs continuously > 5s (PUB006)
 *   - Retention: Held TRUE for mandatory 3s cooldown (PUB006)
 *   - Explicit Reset: Cleared automatically after 3s elapses
 *   - Units: Boolean flag (TRUE = protection latched)
 * -----------------------------------------------------------
 * CurrentTemperature / SetTempDisplay (REAL, output):
 *   - Activation: Assigned every scan from inputs (PUB007)
 *   - Units: degrees
 * -----------------------------------------------------------
 * HeaterStatus (BOOL, output):
 *   - Activation: Mirrors HeaterOutput each scan (PUB007)
 *   - Units: Boolean status indicator
 * ============================================================
 * CONTRACT_RULES []
 * ============================================================ *)

tmp_SensorFault := (TemperatureSensorInput < 0.0) OR (TemperatureSensorInput > 100.0);

CurrentTemperature := TemperatureSensorInput;
SetTempDisplay := SetTemperature;

IF tmp_SensorFault THEN
    HeaterOnRequest := FALSE;
ELSIF OverheatProtection THEN
    HeaterOnRequest := FALSE;
ELSE
    HeaterOnRequest := (TemperatureSensorInput < SetTemperature);
END_IF;

OverheatTimer(IN := HeaterOnRequest AND NOT OverheatProtection,
              PT := T#5S);

IF OverheatTimer.Q THEN
    OverheatProtection := TRUE;
END_IF;

OverheatCooldownTimer(IN := OverheatProtection,
                      PT := T#3S);

IF OverheatCooldownTimer.Q THEN
    OverheatProtection := FALSE;
END_IF;

IF tmp_SensorFault THEN
    HeaterOutput := FALSE;
ELSIF OverheatProtection THEN
    HeaterOutput := FALSE;
ELSE
    HeaterOutput := HeaterOnRequest;
END_IF;

HeaterStatus := HeaterOutput;

END_FUNCTION_BLOCK

(* ---- public-medium-04.candidate_04.st ---- *)
FUNCTION_BLOCK FB_TemperatureControl
VAR_INPUT
    TemperatureSensorInput : REAL;
    SetTemperature : REAL;
END_VAR
VAR_OUTPUT
    CurrentTemperature : REAL;
    SetTempDisplay : REAL;
    HeaterStatus : BOOL;
    OverheatProtection : BOOL;
    HeaterOutput : BOOL;
END_VAR
VAR
    HeaterOnRequest : BOOL;
    tmp_SensorFault : BOOL;
    tmp_AccumulatedHeaterOnTime : LTIME;
    tmp_AccumulatedCooldownTime : LTIME;
END_VAR

(* ENGINEERING_CONTRACT
 * ============================================================
 * Outputs & State Groups:
 * -----------------------------------------------------------
 * HeaterOutput (BOOL, output):
 *   - Activation: Set TRUE when temp < set, no fault, no overheat
 *   - Retention: Maintained TRUE across scans while conditions hold
 *   - Explicit Reset: Set FALSE by fault OR overheat trigger (same-scan)
 *   - Same-scan Priority: OverheatProtection > Fault > Temperature
 *   - Units: Boolean on/off signal
 * -----------------------------------------------------------
 * OverheatProtection (BOOL, output):
 *   - Activation: Set TRUE after heater runs continuously > 5s (PUB006)
 *   - Retention: Held TRUE for mandatory 3s cooldown (PUB006)
 *   - Explicit Reset: Cleared automatically after 3s elapses
 *   - Units: Boolean flag (TRUE = protection latched)
 * -----------------------------------------------------------
 * CurrentTemperature / SetTempDisplay (REAL, output):
 *   - Activation: Assigned every scan from inputs (PUB007)
 *   - Units: degrees
 * -----------------------------------------------------------
 * HeaterStatus (BOOL, output):
 *   - Activation: Mirrors HeaterOutput each scan (PUB007)
 *   - Units: Boolean status indicator
 * ============================================================
 * CONTRACT_RULES []
 * ============================================================ *)

tmp_SensorFault := (TemperatureSensorInput < 0.0) OR (TemperatureSensorInput > 100.0);

CurrentTemperature := TemperatureSensorInput;
SetTempDisplay := SetTemperature;

IF tmp_SensorFault THEN
    HeaterOnRequest := FALSE;
    tmp_AccumulatedHeaterOnTime := LTIME#0s;
ELSIF OverheatProtection THEN
    HeaterOnRequest := FALSE;
ELSE
    HeaterOnRequest := (TemperatureSensorInput < SetTemperature);
END_IF;

IF HeaterOnRequest THEN
    tmp_AccumulatedHeaterOnTime := tmp_AccumulatedHeaterOnTime + TON_Accumulator(HeaterOnRequest);
    IF tmp_AccumulatedHeaterOnTime >= LTIME#5s THEN
        OverheatProtection := TRUE;
        tmp_AccumulatedHeaterOnTime := LTIME#0s;
        HeaterOnRequest := FALSE;
    END_IF;
END_IF;

IF OverheatProtection THEN
    tmp_AccumulatedCooldownTime := tmp_AccumulatedCooldownTime + TON_Accumulator(OverheatProtection);
    IF tmp_AccumulatedCooldownTime >= LTIME#3s THEN
        OverheatProtection := FALSE;
        tmp_AccumulatedCooldownTime := LTIME#0s;
    END_IF;
END_IF;

IF tmp_SensorFault THEN
    HeaterOutput := FALSE;
ELSIF OverheatProtection THEN
    HeaterOutput := FALSE;
ELSE
    HeaterOutput := HeaterOnRequest;
END_IF;

HeaterStatus := HeaterOutput;

END_FUNCTION_BLOCK

(* ---- public-medium-04.raw_candidate_01.st ---- *)
FUNCTION_BLOCK FB_TemperatureControl
VAR_INPUT
    TemperatureSensorInput : REAL;
    SetTemperature : REAL;
END_VAR
VAR_OUTPUT
    CurrentTemperature : REAL;
    SetTempDisplay : REAL;
    HeaterStatus : BOOL;
    OverheatProtection : BOOL;
    HeaterOutput : BOOL;
END_VAR
VAR
    HeaterOnRequest : BOOL;
    OverheatTimer : TON;
    OverheatCooldownTimer : TON;
    tmp_SensorFault : BOOL;
    tmp_HeaterShouldBeOn : BOOL;
END_VAR

(* ENGINEERING_CONTRACT
 * ============================================================
 * Outputs & State Groups:
 * -----------------------------------------------------------
 * HeaterOutput (BOOL, output):
 *   - Activation: Set TRUE when temp < set, no fault, no overheat
 *   - Retention: Maintained TRUE across scans while conditions hold
 *   - Explicit Reset: Set FALSE by fault detection OR overheat trigger
 *   - Same-scan Priority: Fault > Overheat > Temperature comparison
 *   - Units: Boolean on/off signal
 * -----------------------------------------------------------
 * OverheatProtection (BOOL, output):
 *   - Activation: Set TRUE after heater runs continuously > 5s (PUB006)
 *   - Retention: Held TRUE for mandatory 3s cooldown period (PUB006)
 *   - Explicit Reset: Cleared automatically after 3s elapses
 *   - Same-scan Priority: Timer expiry drives reset after 3s
 *   - Units: Boolean flag (TRUE = protection latched)
 * -----------------------------------------------------------
 * CurrentTemperature / SetTempDisplay (REAL, output):
 *   - Activation: Assigned every scan from inputs
 *   - Retention: No retention; mirrors inputs each scan
 *   - Explicit Reset: N/A (always reflects current values)
 *   - Same-scan Priority: Direct assignment
 *   - Units: degrees (temperature values, PUB002/PUB007)
 * -----------------------------------------------------------
 * HeaterStatus (BOOL, output):
 *   - Activation: Mirrors HeaterOutput value each scan
 *   - Retention: Reflects current heater state
 *   - Explicit Reset: Same as HeaterOutput
 *   - Units: Boolean status indicator (PUB007)
 * ============================================================
 * CONTRACT_RULES []
 * ============================================================ *)

tmp_SensorFault := (TemperatureSensorInput < 0.0) OR (TemperatureSensorInput > 100.0);

CurrentTemperature := TemperatureSensorInput;
SetTempDisplay := SetTemperature;

IF tmp_SensorFault THEN
    HeaterOnRequest := FALSE;
ELSIF OverheatProtection THEN
    HeaterOnRequest := FALSE;
ELSE
    tmp_HeaterShouldBeOn := (TemperatureSensorInput < SetTemperature);
    HeaterOnRequest := tmp_HeaterShouldBeOn;
END_IF;

OverheatTimer(IN := HeaterOnRequest AND NOT OverheatProtection,
              PT := T#5S);

IF OverheatTimer.Q THEN
    OverheatProtection := TRUE;
END_IF;

OverheatCooldownTimer(IN := OverheatProtection,
                      PT := T#3S);

IF OverheatCooldownTimer.Q THEN
    OverheatProtection := FALSE;
END_IF;

HeaterOutput := HeaterOnRequest;
HeaterStatus := HeaterOutput;

END_FUNCTION_BLOCK

(* ---- public-medium-04.raw_candidate_02.st ---- *)
FUNCTION_BLOCK FB_TemperatureControl
VAR_INPUT
    TemperatureSensorInput : REAL;
    SetTemperature : REAL;
END_VAR
VAR_OUTPUT
    CurrentTemperature : REAL;
    SetTempDisplay : REAL;
    HeaterStatus : BOOL;
    OverheatProtection : BOOL;
    HeaterOutput : BOOL;
END_VAR
VAR
    HeaterOnRequest : BOOL;
    OverheatTimer : TON;
    CooldownTimer : TON;
    tmp_SensorFault : BOOL;
    tmp_HeaterShouldBeOn : BOOL;
END_VAR

(* ENGINEERING_CONTRACT
 * ============================================================
 * Outputs & State Groups:
 * -----------------------------------------------------------
 * HeaterOutput (BOOL, output):
 *   - Activation: Set TRUE when temp < set, no fault, no overheat
 *   - Retention: Maintained TRUE across scans while conditions hold
 *   - Explicit Reset: Set FALSE by fault detection OR overheat trigger
 *   - Same-scan Priority: Fault > Overheat > Temperature comparison
 *   - Units: Boolean on/off signal
 * -----------------------------------------------------------
 * OverheatProtection (BOOL, output):
 *   - Activation: Set TRUE after heater runs continuously > 5s (PUB006)
 *   - Retention: Held TRUE for mandatory 3s cooldown period (PUB006)
 *   - Explicit Reset: Cleared automatically after 3s elapses
 *   - Same-scan Priority: Timer expiry drives reset after 3s
 *   - Units: Boolean flag (TRUE = protection latched)
 * -----------------------------------------------------------
 * CurrentTemperature / SetTempDisplay (REAL, output):
 *   - Activation: Assigned every scan from inputs
 *   - Retention: No retention; mirrors inputs each scan
 *   - Explicit Reset: N/A (always reflects current values)
 *   - Units: degrees (temperature values, PUB002/PUB007)
 * -----------------------------------------------------------
 * HeaterStatus (BOOL, output):
 *   - Activation: Mirrors HeaterOutput value each scan
 *   - Retention: Reflects current heater state
 *   - Units: Boolean status indicator (PUB007)
 * ============================================================
 * CONTRACT_RULES []
 * ============================================================ *)

tmp_SensorFault := (TemperatureSensorInput < 0.0) OR (TemperatureSensorInput > 100.0);

CurrentTemperature := TemperatureSensorInput;
SetTempDisplay := SetTemperature;

IF tmp_SensorFault THEN
    HeaterOnRequest := FALSE;
ELSIF OverheatProtection THEN
    HeaterOnRequest := FALSE;
ELSE
    tmp_HeaterShouldBeOn := (TemperatureSensorInput < SetTemperature);
    HeaterOnRequest := tmp_HeaterShouldBeOn;
END_IF;

OverheatTimer(IN := HeaterOnRequest AND NOT OverheatProtection,
              PT := T#5S);

IF OverheatTimer.Q THEN
    OverheatProtection := TRUE;
END_IF;

CooldownTimer(IN := OverheatProtection,
              PT := T#3S);

IF CooldownTimer.Q THEN
    OverheatProtection := FALSE;
END_IF;

HeaterOutput := HeaterOnRequest;
HeaterStatus := HeaterOutput;

END_FUNCTION_BLOCK

(* ---- public-medium-04.raw_candidate_03.st ---- *)
FUNCTION_BLOCK FB_TemperatureControl
VAR_INPUT
    TemperatureSensorInput : REAL;
    SetTemperature : REAL;
END_VAR
VAR_OUTPUT
    CurrentTemperature : REAL;
    SetTempDisplay : REAL;
    HeaterStatus : BOOL;
    OverheatProtection : BOOL;
    HeaterOutput : BOOL;
END_VAR
VAR
    HeaterOnRequest : BOOL;
    OverheatTimer : TON;
    OverheatCooldownTimer : TON;
    tmp_SensorFault : BOOL;
END_VAR

(* ENGINEERING_CONTRACT
 * ============================================================
 * Outputs & State Groups:
 * -----------------------------------------------------------
 * HeaterOutput (BOOL, output):
 *   - Activation: Set TRUE when temp < set, no fault, no overheat
 *   - Retention: Maintained TRUE across scans while conditions hold
 *   - Explicit Reset: Set FALSE by fault OR overheat trigger (same-scan)
 *   - Same-scan Priority: OverheatProtection > Fault > Temperature
 *   - Units: Boolean on/off signal
 * -----------------------------------------------------------
 * OverheatProtection (BOOL, output):
 *   - Activation: Set TRUE after heater runs continuously > 5s (PUB006)
 *   - Retention: Held TRUE for mandatory 3s cooldown (PUB006)
 *   - Explicit Reset: Cleared automatically after 3s elapses
 *   - Units: Boolean flag (TRUE = protection latched)
 * -----------------------------------------------------------
 * CurrentTemperature / SetTempDisplay (REAL, output):
 *   - Activation: Assigned every scan from inputs (PUB007)
 *   - Units: degrees
 * -----------------------------------------------------------
 * HeaterStatus (BOOL, output):
 *   - Activation: Mirrors HeaterOutput each scan (PUB007)
 *   - Units: Boolean status indicator
 * ============================================================
 * CONTRACT_RULES []
 * ============================================================ *)

tmp_SensorFault := (TemperatureSensorInput < 0.0) OR (TemperatureSensorInput > 100.0);

CurrentTemperature := TemperatureSensorInput;
SetTempDisplay := SetTemperature;

IF tmp_SensorFault THEN
    HeaterOnRequest := FALSE;
ELSIF OverheatProtection THEN
    HeaterOnRequest := FALSE;
ELSE
    HeaterOnRequest := (TemperatureSensorInput < SetTemperature);
END_IF;

OverheatTimer(IN := HeaterOnRequest AND NOT OverheatProtection,
              PT := T#5S);

IF OverheatTimer.Q THEN
    OverheatProtection := TRUE;
END_IF;

OverheatCooldownTimer(IN := OverheatProtection,
                      PT := T#3S);

IF OverheatCooldownTimer.Q THEN
    OverheatProtection := FALSE;
END_IF;

IF tmp_SensorFault THEN
    HeaterOutput := FALSE;
ELSIF OverheatProtection THEN
    HeaterOutput := FALSE;
ELSE
    HeaterOutput := HeaterOnRequest;
END_IF;

HeaterStatus := HeaterOutput;

END_FUNCTION_BLOCK
